// Mitsubishi GX Works2 project: Cascade3_V4   PLC: FX3G

TYPE PUMP : STRUCT
  Blocked : BOOL;
  Start : BOOL;
  Evailable : BOOL;
END_STRUCT END_TYPE

TYPE BURNER : STRUCT
  Manual : BOOL;
  Auto : BOOL;
  Stage1 : BOOL;
  Stage2 : BOOL;
  Pressure : INT;
  Temperature : INT;
  Power : BOOL;
  Work : BOOL;
  ManualSecond : BOOL;  (* Назначить горелку на вторую ступень *)
  Error : BOOL;
  Enable : BOOL;
END_STRUCT END_TYPE

// global labels: IO
VAR_GLOBAL
  AI_T_Heater1 AT D0 : INT;  (* Температура котла №1 с модуля АЦП (R23700), °C x10 *)
  AI_T_Heater2 AT D1 : INT;  (* Температура котла №2 с модуля АЦП (R23701), °C x10 *)
  AI_T_Heater3 AT D2 : INT;  (* Температура котла №3 с модуля АЦП (R23702), °C x10 *)
  AI_T_Colector AT D3 : INT;  (* Температура обратки с коллектора (R23703), °C x10 *)
  AI_T_SOFrom AT D4 : INT;  (* Температура обратки отопления (R23704), °C x10 *)
  AI_T_SOTo AT D5 : INT;  (* Температура подачи отопления (R23705), °C x10 *)
  AI_T_GVSTo AT D6 : INT;  (* Температура подачи на теплообменник ГВС (R23706), °C x10 *)
  AI_T_GVSFrom AT D7 : INT;  (* Температура обратки с теплообменника ГВС (R23707), °C x10 *)
  AI_T_Gaz AT D8 : INT;  (* Температура газа (R23709), °C x10 *)
  AI_T_Weather AT D9 : INT;  (* Температура наружного воздуха (R23708), °C x10 *)
  AI_P1 AT D10 : INT;  (* Давление в котле №1 с датчика, в десятых долях (шкала задаётся в Max_P1) *)
  AI_P2 AT D11 : INT;  (* Давление в котле №2 с датчика, в десятых долях (шкала задаётся в Max_P2) *)
  AI_P3 AT D12 : INT;  (* Давление в котле №3 с датчика, в десятых долях (шкала задаётся в Max_P3) *)
  AI_P_SOTo AT D13 : INT;  (* Давление подачи отопления с датчика, в десятых долях (шкала задаётся в Max_P_SOTo) *)
  AI_P_SOFrom AT D14 : INT;  (* Давление обратки отопления с датчика, в десятых долях (шкала задаётся в Max_P_SOFrom) *)
  AI_P_GVSTo AT D15 : INT;  (* Давление подачи на теплообменник с датчика, в десятых долях (шкала задаётся в Max_P_GVSTo) *)
  AI_P_GVSFrom AT D16 : INT;  (* Давление обратки с теплообменника с датчика, в десятых долях (шкала задаётся в Max_P_GVSFrom) *)
  AI_P_Set AT D17 : INT;  (* Давление в системе (подпитка), в десятых долях. D35 занят, поэтому D17 *)
  AI_P_GAZ AT D18 : INT;  (* Давление газа с датчика (D8032), в десятых долях *)
  DI_EKM AT X000 : BOOL;  (* Реле давления (ЭКМ): контакт разомкнут — авария 26 *)
  DI_ES AT X001 : BOOL;  (* Кнопка аварийного отключения: снимает gxStart, авария 27 *)
  DI_RKF AT X010 : BOOL;  (* Реле контроля фаз: контакт разомкнут — авария 28 *)
  DI_BurnAlarm1 AT X002 : BOOL;  (* Сухой контакт «авария горелки №1» *)
  DI_BurnAlarm2 AT X003 : BOOL;  (* Сухой контакт «авария горелки №2» *)
  DI_BurnAlarm3 AT X004 : BOOL;  (* Сухой контакт «авария горелки №3» *)
  DI_BurnWork1 AT X005 : BOOL;  (* Сухой контакт «горелка №1 в работе» *)
  DI_BurnWork2 AT X006 : BOOL;  (* Сухой контакт «горелка №2 в работе» *)
  DI_BurnWork3 AT X007 : BOOL;  (* Сухой контакт «горелка №3 в работе» *)
  DI_Pump1_T1 AT X011 : BOOL;  (* Обратная связь: насос №1 контура Т1 работает *)
  DI_Pump2_T1 AT X012 : BOOL;  (* Обратная связь: насос №2 контура Т1 работает *)
  DI_Pump1_T1_2 AT X013 : BOOL;  (* Обратная связь: насос №1 контура Т1.2 работает *)
  DI_Pump2_T1_2 AT X020 : BOOL;  (* Обратная связь: насос №2 контура Т1.2 работает *)
  DI_Pump1_T3 AT X021 : BOOL;  (* Обратная связь: насос №1 контура Т3 работает *)
  DI_Pump2_T3 AT X022 : BOOL;  (* Обратная связь: насос №2 контура Т3 работает *)
  DI_Pump1 AT X023 : BOOL;  (* Обратная связь: насос циркуляции №1 малого контура работает *)
  DI_Pump2 AT X024 : BOOL;  (* Обратная связь: насос циркуляции №2 малого контура работает *)
  DI_Pump3 AT X025 : BOOL;  (* Обратная связь: насос циркуляции №3 малого контура работает *)
  DI_AlarmReset AT X030 : BOOL;  (* Внешняя кнопка сброса аварий и сирены *)
  DI_BurnTherm1 AT X035 : BOOL;  (* Термозащита котла №1: нормально замкнутый контакт, нет цепи — авария *)
  DI_BurnTherm2 AT X036 : BOOL;  (* Термозащита котла №2: нормально замкнутый контакт, нет цепи — авария *)
  DI_BurnTherm3 AT X037 : BOOL;  (* Термозащита котла №3: нормально замкнутый контакт, нет цепи — авария *)
  DO_Burn1Power AT Y035 : BOOL;  (* Разрешение работы (питание) горелки №1: без него ступени не включаются *)
  DO_Burn1Stage1 AT Y000 : BOOL;  (* Горелка №1: включить ступень 1 *)
  DO_Burn1Stage2 AT Y001 : BOOL;  (* Горелка №1: включить ступень 2 *)
  DO_Burn2Power AT Y036 : BOOL;  (* Разрешение работы (питание) горелки №2: без него ступени не включаются *)
  DO_Burn2Stage1 AT Y002 : BOOL;  (* Горелка №2: включить ступень 1 *)
  DO_Burn2Stage2 AT Y003 : BOOL;  (* Горелка №2: включить ступень 2 *)
  DO_Burn3Power AT Y037 : BOOL;  (* Разрешение работы (питание) горелки №3: без него ступени не включаются *)
  DO_Burn3Stage1 AT Y004 : BOOL;  (* Горелка №3: включить ступень 1 *)
  DO_Burn3Stage2 AT Y005 : BOOL;  (* Горелка №3: включить ступень 2 *)
  DO_ValveFill AT Y006 : BOOL;  (* Клапан набора воды (подпитка) *)
  DO_AlarmBuzzer AT Y007 : BOOL;  (* Сирена: звуковая сигнализация аварии *)
  DO_AlarmLight AT Y010 : BOOL;  (* Лампа аварии *)
  DO_Pump1_T1 AT Y020 : BOOL;  (* Включить насос №1 контура Т1 *)
  DO_Pump2_T1 AT Y021 : BOOL;  (* Включить насос №2 контура Т1 *)
  DO_Pump1_T1_2 AT Y022 : BOOL;  (* Включить насос №1 контура Т1.2 *)
  DO_Pump2_T1_2 AT Y023 : BOOL;  (* Включить насос №2 контура Т1.2 *)
  DO_Pump1_T3 AT Y024 : BOOL;  (* Включить насос №1 контура Т3 *)
  DO_Pump2_T3 AT Y025 : BOOL;  (* Включить насос №2 контура Т3 *)
  DO_Pump1 AT Y026 : BOOL;  (* Включить насос циркуляции №1 малого контура *)
  DO_Pump2 AT Y027 : BOOL;  (* Включить насос циркуляции №2 малого контура *)
  DO_Pump3 AT Y030 : BOOL;  (* Включить насос циркуляции №3 малого контура *)
  DO_3wayOpen AT Y033 : BOOL;  (* 3-ходовой клапан: открыть *)
  DO_3wayClose AT Y034 : BOOL;  (* 3-ходовой клапан: закрыть *)
END_VAR

// global labels: GVL
VAR_GLOBAL
  arBurners : ARRAY [0..2] OF BURNER;  (* (Set M500) Состояние трёх котлов (структура BURNER): включён в авто, ступень 1, ступень 2, авария, ручной режим *)
END_VAR
VAR_GLOBAL CONSTANT
  c_HEATERS : INT := 3;  (* Количество котлов в каскаде *)
  c_HEATERS_IDX : INT := 2;  (* Индекс последнего котла в массиве (c_HEATERS - 1) *)
  c_AM_ALARMS_NUM : INT := 54;  (* Верхняя граница массива аварий: используются номера 0…45 (46 штук). Максимум 127 *)
END_VAR
VAR_GLOBAL
  AM_ALARMS : ARRAY [0..54] OF ST_AM_ALARM;  (* Массив аварий менеджера тревог. Граница 45 должна совпадать с c_AM_ALARMS_NUM. Состояние: AM_ALARMS[i].Alarm *)
  gxStart AT M400 : BOOL;  (* Пуск/останов каскада с панели (1 = работа). Снимается кнопкой X001 и авариями *)
  gxErrorReset AT M401 : BOOL;  (* Сброс всех аварий (1 = сбросить). В шаге 0 выставляется программой автоматически *)
  gxHasalarm AT M402 : BOOL;  (* Есть хотя бы одна активная авария. Формируется блоком FB_AM_HAS_ALARMS, используется для лампы и панели *)
  gxNoSettings AT M403 : BOOL;  (* Не заданы уставки или коэффициенты ПИД (R503 = 0). Пуск запрещён, авария 30 *)
  gxResetAlarm AT M404 : BOOL;  (* Кнопка «Сброс сигнализации» на панели: снимает сирену и лампу *)
  gxFillManual AT M405 : BOOL;  (* Ручной режим подпитки: клапан набора воды открыт, пока флаг включён *)
  gxFillAuto AT M406 : BOOL;  (* Автоматическая подпитка по давлению в системе (SV_PresFilStart / SV_PresFilStop) *)
  gxResetWHT1 AT M407 : BOOL;  (* Сброс моточасов котла №1 (giHeater1Hours) *)
  gxResetWHT2 AT M408 : BOOL;  (* Сброс моточасов котла №2 (giHeater2Hours) *)
  gxResetWHT3 AT M409 : BOOL;  (* Сброс моточасов котла №3 (giHeater3Hours) *)
  gxPIDAT AT M410 : BOOL;  (* Запуск автонастройки ПИД каскада (блок параметров R500…R528). Сбрасывается сама по завершении *)
  gxPIDATLimitCycle AT M411 : BOOL;  (* Ограничение числа циклов автонастройки ПИД каскада: 0 — не больше 50, 1 — не больше 114 *)
  gxEnablePump1 AT M412 : BOOL;  (* Разрешение насоса циркуляции №1 малого контура (1 = участвует в работе) *)
  gxEnablePump2 AT M413 : BOOL;  (* Разрешение насоса циркуляции №2 малого контура (1 = участвует в работе) *)
  gxEnablePump3 AT M415 : BOOL;  (* Разрешение насоса циркуляции №3 малого контура (1 = участвует в работе). M414 пропущен — так привязано на панели *)
  gxManualPump1 AT M416 : BOOL;  (* Ручной пуск насоса циркуляции №1 малого контура (нужно ещё разрешение gxEnablePump1) *)
  gxManualPump2 AT M417 : BOOL;  (* Ручной пуск насоса циркуляции №2 малого контура (нужно ещё разрешение gxEnablePump2) *)
  gxManualPump3 AT M418 : BOOL;  (* Ручной пуск насоса циркуляции №3 малого контура (нужно ещё разрешение gxEnablePump3) *)
  gx3WayCloseWhenOff AT M419 : BOOL;  (* Закрывать 3-ходовой клапан при останове каскада (1 = закрывать) *)
  gxPID3WayAT AT M420 : BOOL;  (* Запуск автонастройки ПИД 3-ходового клапана (блок параметров R600…R628) *)
  gxPID3WayATLimitCycle AT M421 : BOOL;  (* Ограничение числа циклов автонастройки ПИД 3-ходового клапана: 0 — не больше 50, 1 — не больше 114 *)
  gxPump1_T1_Enable AT M422 : BOOL;  (* Разрешение насоса №1 контура Т1 (1 = участвует в каскаде, 0 = заблокирован) *)
  gxPump2_T1_Enable AT M423 : BOOL;  (* Разрешение насоса №2 контура Т1 (1 = участвует в каскаде, 0 = заблокирован) *)
  gxPump1_T1_2_Enable AT M424 : BOOL;  (* Разрешение насоса №1 контура Т1.2 (1 = участвует в каскаде, 0 = заблокирован) *)
  gxPump2_T1_2_Enable AT M425 : BOOL;  (* Разрешение насоса №2 контура Т1.2 (1 = участвует в каскаде, 0 = заблокирован) *)
  gxPump1_T3_Enable AT M426 : BOOL;  (* Разрешение насоса №1 контура Т3 (1 = участвует в каскаде, 0 = заблокирован) *)
  gxPump2_T3_Enable AT M427 : BOOL;  (* Разрешение насоса №2 контура Т3 (1 = участвует в каскаде, 0 = заблокирован) *)
  gxPump1_T1_Manual AT M428 : BOOL;  (* Ручной пуск насоса №1 контура Т1 *)
  gxPump2_T1_Manual AT M429 : BOOL;  (* Ручной пуск насоса №2 контура Т1 *)
  gxPump1_T1_2_Manual AT M430 : BOOL;  (* Ручной пуск насоса №1 контура Т1.2 *)
  gxPump2_T1_2_Manual AT M431 : BOOL;  (* Ручной пуск насоса №2 контура Т1.2 *)
  gxPump1_T3_Manual AT M432 : BOOL;  (* Ручной пуск насоса №1 контура Т3 *)
  gxPump2_T3_Manual AT M433 : BOOL;  (* Ручной пуск насоса №2 контура Т3 *)
  gxPump1_T1_WHReset AT M434 : BOOL;  (* Сброс моточасов насоса №1 контура Т1 *)
  gxPump2_T1_WHReset AT M435 : BOOL;  (* Сброс моточасов насоса №2 контура Т1 *)
  gxPump1_T1_2_WHReset AT M436 : BOOL;  (* Сброс моточасов насоса №1 контура Т1.2 *)
  gxPump2_T1_2_WHReset AT M437 : BOOL;  (* Сброс моточасов насоса №2 контура Т1.2 *)
  gxPump1_T3_WHReset AT M438 : BOOL;  (* Сброс моточасов насоса №1 контура Т3 *)
  gxPump2_T3_WHReset AT M439 : BOOL;  (* Сброс моточасов насоса №2 контура Т3 *)
  gxPump1_WHReset AT M440 : BOOL;  (* Сброс моточасов насоса циркуляции №1 малого контура *)
  gxPump2_WHReset AT M441 : BOOL;  (* Сброс моточасов насоса циркуляции №2 малого контура *)
  gxPump3_WHReset AT M442 : BOOL;  (* Сброс моточасов насоса циркуляции №3 малого контура *)
  gx3WayEnable AT M443 : BOOL;  (* Разрешение работы 3-ходового клапана (1 = регулирует, 0 = стоит) *)
  gx3WayManual AT M444 : BOOL;  (* Ручной режим 3-ходового клапана: положение берётся из SV_3WayManualTask, ПИД отключён *)
  gxWHOvfHeater1 AT M450 : BOOL;  (* Переполнение счётчика моточасов котла №1 (выход HOUR). 1 — счётчик переполнен, нужно сбросить *)
  gxWHOvfHeater2 AT M451 : BOOL;  (* Переполнение счётчика моточасов котла №2 (выход HOUR). 1 — счётчик переполнен, нужно сбросить *)
  gxWHOvfHeater3 AT M452 : BOOL;  (* Переполнение счётчика моточасов котла №3 (выход HOUR). 1 — счётчик переполнен, нужно сбросить *)
  gxWHOvfPump1_T1 AT M453 : BOOL;  (* Переполнение счётчика моточасов насоса №1 контура Т1 (выход HOUR) *)
  gxWHOvfPump2_T1 AT M454 : BOOL;  (* Переполнение счётчика моточасов насоса №2 контура Т1 (выход HOUR) *)
  gxWHOvfPump1_T1_2 AT M455 : BOOL;  (* Переполнение счётчика моточасов насоса №1 контура Т1.2 (выход HOUR) *)
  gxWHOvfPump2_T1_2 AT M456 : BOOL;  (* Переполнение счётчика моточасов насоса №2 контура Т1.2 (выход HOUR) *)
  gxWHOvfPump1_T3 AT M457 : BOOL;  (* Переполнение счётчика моточасов насоса №1 контура Т3 (выход HOUR) *)
  gxWHOvfPump2_T3 AT M458 : BOOL;  (* Переполнение счётчика моточасов насоса №2 контура Т3 (выход HOUR) *)
  gxWHOvfPump1 AT M459 : BOOL;  (* Переполнение счётчика моточасов насоса циркуляции №1 (выход HOUR) *)
  gxWHOvfPump2 AT M460 : BOOL;  (* Переполнение счётчика моточасов насоса циркуляции №2 (выход HOUR) *)
  gxWHOvfPump3 AT M461 : BOOL;  (* Переполнение счётчика моточасов насоса циркуляции №3 (выход HOUR) *)
  giPIDTask AT D500 : INT;  (* Выход ПИД каскада: задание в ступенях мощности (0…6). Из него считается, сколько котлов и ступеней включить *)
  giTSV AT D501 : INT;  (* Текущее задание температуры теплоносителя: по кривой погодозависимости или SV_TWater1, если на улице тепло *)
  giAvailableStages AT D502 : INT;  (* Сколько ступеней доступно автоматике: по 2 на каждый котёл в авто без аварий *)
  giWorkStages AT D503 : INT;  (* Сколько ступеней включено сейчас в авторежиме *)
  giPID3WayTask AT D504 : INT;  (* Выход ПИД 3-ходового клапана: положение 0…1000 (0.0…100.0 %, 0 — закрыт, 1000 — открыт). Диапазон задан R622 = 1000 *)
  SV_3WayTempGVS AT D510 : INT;  (* Уставка температуры ГВС на выходе теплообменника, °C *)
  SV_MaxTemperatureHeater AT D511 : INT;  (* Максимальная температура котла, °C. Выше — авария перегрева *)
  SV_TLimit AT D512 : INT;  (* Допустимое превышение задания, °C: котёл отключается при температуре выше задания на эту величину *)
  SV_HowOftenToCheck AT D513 : INT;  (* Как часто проверять каскад (добавлять или убирать ступени), секунд *)
  SV_MaxPressure AT D514 : INT;  (* Максимальное давление в котле (авария). В тех же единицах, что и показания датчика *)
  SV_MinPressure AT D515 : INT;  (* Минимальное давление в котле (авария) *)
  SV_PresFilStart AT D516 : INT;  (* Давление в системе, при котором начинается подпитка *)
  SV_PresFilStop AT D517 : INT;  (* Давление в системе, при котором подпитка заканчивается *)
  SV_GasMinPressure AT D518 : INT;  (* Минимальное давление газа. Ниже — авария 24 и блокировка каскада *)
  SV_SetMinPressure AT D519 : INT;  (* Минимальное давление в системе. Ниже — авария 25 и запрет циркуляционных насосов *)
  SV_MaxFillTime AT D520 : INT;  (* Максимальное время набора воды, секунд. Дольше — авария 34 *)
  SV_TimeinWork AT D521 : INT;  (* Резерв: в программе не используется (осталось от старой версии), выводится только на панель *)
  SV_3WayDelta AT D522 : INT;  (* Зона нечувствительности 3-ходового клапана в единицах положения 0…1000 (50 = 5.0 %); в ручном режиме принудительно равна 0 *)
  SV_3WayTotalTime AT D523 : INT;  (* Полное время хода 3-ходового клапана, секунд *)
  SV_3WayLuftTime AT D524 : INT;  (* Время люфта (мёртвого хода) 3-ходового клапана, миллисекунд *)
  SV_3WayTempGVSDelta AT D525 : INT;  (* Гистерезис по ГВС, °C: ПИД работает, пока температура ниже уставки на эту величину *)
  SV_3WayManualTask AT D526 : INT;  (* Задание положения 3-ходового клапана в ручном режиме, 0…1000 (0.1 % за единицу) — та же шкала, что у выхода ПИД *)
  SV_3WayMaxTemperature AT D527 : INT;  (* Максимальная температура ГВС, °C. Выше — авария 35 *)
  SV_MaxTemperatureColector AT D528 : INT;  (* Максимальная температура коллектора, °C. Выше — авария 32 и отключение ПИД каскада *)
  SV_StageHyst AT D583 : INT;  (* % x10 с панели (50 = 5.0 %). Зона нечувствительности добавления ступени: насколько выход ПИД (0…600 = 0…100 %) должен превысить границу следующей ступени, чтобы включилась ещё одна ступень. Убираются ступени без задержки. ПЛК пересчитывает проценты в единицы ПИД: iHyst = значение * 6 / 10 *)
  giHeater1Hours AT D560 : ARRAY [0..1] OF INT;  (* Наработка котла №1, моточасы (массив из 2 слов для счётчика HOUR) *)
  giHeater2Hours AT D562 : ARRAY [0..1] OF INT;  (* Наработка котла №2, моточасы (массив из 2 слов для счётчика HOUR) *)
  giHeater3Hours AT D564 : ARRAY [0..1] OF INT;  (* Наработка котла №3, моточасы (массив из 2 слов для счётчика HOUR) *)
  T1_State AT D566 : INT;  (* Состояние котла №1 для панели: 0 — не разрешён, 1 — разрешён и стоит, 2 — ступень 1, 3 — ступень 2 *)
  T2_State AT D567 : INT;  (* Состояние котла №2 для панели: 0 — не разрешён, 1 — разрешён и стоит, 2 — ступень 1, 3 — ступень 2 *)
  T3_State AT D568 : INT;  (* Состояние котла №3 для панели: 0 — не разрешён, 1 — разрешён и стоит, 2 — ступень 1, 3 — ступень 2 *)
  Pump1_T1_State AT D569 : INT;  (* Состояние насоса №1 контура Т1 для панели: 0 — стоит, 1 — работает, 2 — авария, 4 — заблокирован *)
  Pump2_T1_State AT D570 : INT;  (* Состояние насоса №2 контура Т1 для панели: 0 — стоит, 1 — работает, 2 — авария, 4 — заблокирован *)
  Pump1_T1_2_State AT D571 : INT;  (* Состояние насоса №1 контура Т1.2 для панели: 0 — стоит, 1 — работает, 2 — авария, 4 — заблокирован *)
  Pump2_T1_2_State AT D572 : INT;  (* Состояние насоса №2 контура Т1.2 для панели: 0 — стоит, 1 — работает, 2 — авария, 4 — заблокирован *)
  Pump1_T3_State AT D573 : INT;  (* Состояние насоса №1 контура Т3 для панели: 0 — стоит, 1 — работает, 2 — авария, 4 — заблокирован *)
  Pump2_T3_State AT D574 : INT;  (* Состояние насоса №2 контура Т3 для панели: 0 — стоит, 1 — работает, 2 — авария, 4 — заблокирован *)
  Pump1_State AT D575 : INT;  (* Состояние насоса циркуляции №1 для панели: 0 — стоит, 1 — работает, 2 — авария, 4 — заблокирован *)
  Pump2_State AT D576 : INT;  (* Состояние насоса циркуляции №2 для панели: 0 — стоит, 1 — работает, 2 — авария, 4 — заблокирован *)
  Pump3_State AT D577 : INT;  (* Состояние насоса циркуляции №3 для панели: 0 — стоит, 1 — работает, 2 — авария, 4 — заблокирован *)
  Pump1_T1_WH AT D600 : ARRAY [0..1] OF INT;  (* Моточасы насоса №1 контура Т1 (2 слова, счётчик HOUR). Область D600…D617 не пересекается с состояниями *)
  Pump2_T1_WH AT D602 : ARRAY [0..1] OF INT;  (* Моточасы насоса №2 контура Т1 (2 слова, счётчик HOUR). Область D600…D617 не пересекается с состояниями *)
  Pump1_T1_2_WH AT D604 : ARRAY [0..1] OF INT;  (* Моточасы насоса №1 контура Т1.2 (2 слова, счётчик HOUR). Область D600…D617 не пересекается с состояниями *)
  Pump2_T1_2_WH AT D606 : ARRAY [0..1] OF INT;  (* Моточасы насоса №2 контура Т1.2 (2 слова, счётчик HOUR). Область D600…D617 не пересекается с состояниями *)
  Pump1_T3_WH AT D608 : ARRAY [0..1] OF INT;  (* Моточасы насоса №1 контура Т3 (2 слова, счётчик HOUR). Область D600…D617 не пересекается с состояниями *)
  Pump2_T3_WH AT D610 : ARRAY [0..1] OF INT;  (* Моточасы насоса №2 контура Т3 (2 слова, счётчик HOUR). Область D600…D617 не пересекается с состояниями *)
  Pump1_WH AT D612 : ARRAY [0..1] OF INT;  (* Моточасы насоса циркуляции №1 (2 слова, счётчик HOUR). Область D600…D617 не пересекается с состояниями *)
  Pump2_WH AT D614 : ARRAY [0..1] OF INT;  (* Моточасы насоса циркуляции №2 (2 слова, счётчик HOUR). Область D600…D617 не пересекается с состояниями *)
  Pump3_WH AT D616 : ARRAY [0..1] OF INT;  (* Моточасы насоса циркуляции №3 (2 слова, счётчик HOUR). Область D600…D617 не пересекается с состояниями *)
  SV_TWeather1 AT D530 : INT;  (* Кривая погодозависимости, точка 1: температура на улице, °C *)
  SV_TWater1 AT D531 : INT;  (* Кривая погодозависимости, точка 1: температура подачи в систему, °C *)
  SV_TWeather2 AT D532 : INT;  (* Кривая погодозависимости, точка 2: температура на улице, °C *)
  SV_TWater2 AT D533 : INT;  (* Кривая погодозависимости, точка 2: температура подачи в систему, °C *)
  SV_TWeather3 AT D534 : INT;  (* Кривая погодозависимости, точка 3: температура на улице, °C *)
  SV_TWater3 AT D535 : INT;  (* Кривая погодозависимости, точка 3: температура подачи в систему, °C *)
  SV_TWeather4 AT D536 : INT;  (* Кривая погодозависимости, точка 4: температура на улице, °C *)
  SV_TWater4 AT D537 : INT;  (* Кривая погодозависимости, точка 4: температура подачи в систему, °C *)
  Cor_T_Heater1 AT D540 : INT;  (* Поправка датчика температуры котла №1: прибавляется к показанию, °C x10 *)
  Cor_T_Heater2 AT D541 : INT;  (* Поправка датчика температуры котла №2: прибавляется к показанию, °C x10 *)
  Cor_T_Heater3 AT D542 : INT;  (* Поправка датчика температуры котла №3: прибавляется к показанию, °C x10 *)
  Cor_T_Colector AT D543 : INT;  (* Поправка датчика температуры коллектора: прибавляется к показанию, °C x10 *)
  Cor_T_SOFrom AT D544 : INT;  (* Поправка датчика температуры обратки отопления: прибавляется к показанию, °C x10 *)
  Cor_T_SOTo AT D545 : INT;  (* Поправка датчика температуры подачи отопления: прибавляется к показанию, °C x10 *)
  Cor_T_GVSTo AT D546 : INT;  (* Поправка датчика температуры подачи на теплообменник ГВС: прибавляется к показанию, °C x10 *)
  Cor_T_GVSFrom AT D547 : INT;  (* Поправка датчика температуры обратки с теплообменника ГВС: прибавляется к показанию, °C x10 *)
  Cor_T_Gaz AT D548 : INT;  (* Поправка датчика температуры датчика газа: прибавляется к показанию, °C x10 *)
  Cor_T_Weather AT D549 : INT;  (* Поправка датчика температуры датчика наружной температуры: прибавляется к показанию, °C x10 *)
  Max_P1 AT D550 : INT;  (* Верхний предел шкалы датчика давления котла №1, в десятых долях (160 = 16.0). 0 — не задан *)
  Max_P2 AT D551 : INT;  (* Верхний предел шкалы датчика давления котла №2, в десятых долях (160 = 16.0). 0 — не задан *)
  Max_P3 AT D552 : INT;  (* Верхний предел шкалы датчика давления котла №3, в десятых долях (160 = 16.0). 0 — не задан *)
  Max_P_SOTo AT D553 : INT;  (* Верхний предел шкалы датчика давления подачи отопления, в десятых долях (160 = 16.0). 0 — не задан *)
  Max_P_SOFrom AT D554 : INT;  (* Верхний предел шкалы датчика давления обратки отопления, в десятых долях (160 = 16.0). 0 — не задан *)
  Max_P_GVSTo AT D555 : INT;  (* Верхний предел шкалы датчика давления подачи на теплообменник, в десятых долях (160 = 16.0). 0 — не задан *)
  Max_P_GVSFrom AT D556 : INT;  (* Верхний предел шкалы датчика давления обратки с теплообменника, в десятых долях (160 = 16.0). 0 — не задан *)
  Max_P_Set AT D557 : INT;  (* Верхний предел шкалы датчика давления в системе, в десятых долях (160 = 16.0). 0 — не задан *)
  Max_P_GAZ AT D558 : INT;  (* Верхний предел шкалы датчика давления газа, в десятых долях (160 = 16.0). 0 — не задан *)
  FAI_T_Heater1 AT D20 : REAL;  (* Температура котла №1, °C в реальных единицах (для панели и графиков) *)
  FAI_T_Heater2 AT D22 : REAL;  (* Температура котла №2, °C в реальных единицах (для панели и графиков) *)
  FAI_T_Heater3 AT D24 : REAL;  (* Температура котла №3, °C в реальных единицах (для панели и графиков) *)
  FAI_T_Colector AT D26 : REAL;  (* Температура обратки с коллектора, °C в реальных единицах (для панели и графиков) *)
  FAI_T_SOFrom AT D28 : REAL;  (* Температура обратки отопления, °C в реальных единицах (для панели и графиков) *)
  FAI_T_SOTo AT D30 : REAL;  (* Температура подачи отопления, °C в реальных единицах (для панели и графиков) *)
  FAI_T_GVSTo AT D32 : REAL;  (* Температура подачи на теплообменник ГВС, °C в реальных единицах (для панели и графиков) *)
  FAI_T_GVSFrom AT D34 : REAL;  (* Температура обратки с теплообменника ГВС, °C в реальных единицах (для панели и графиков) *)
  FAI_T_Gaz AT D36 : REAL;  (* Температура газа, °C в реальных единицах (для панели и графиков) *)
  FAI_T_Weather AT D38 : REAL;  (* Температура наружного воздуха, °C в реальных единицах (для панели и графиков) *)
  FAI_P1 AT D40 : REAL;  (* Давление в котле №1 в реальных единицах (для панели и графиков) *)
  FAI_P2 AT D42 : REAL;  (* Давление в котле №2 в реальных единицах (для панели и графиков) *)
  FAI_P3 AT D44 : REAL;  (* Давление в котле №3 в реальных единицах (для панели и графиков) *)
  FAI_P_SOTo AT D46 : REAL;  (* Давление подачи отопления в реальных единицах (для панели и графиков) *)
  FAI_P_SOFrom AT D48 : REAL;  (* Давление обратки отопления в реальных единицах (для панели и графиков) *)
  FAI_P_GVSTo AT D50 : REAL;  (* Давление подачи на теплообменник в реальных единицах (для панели и графиков) *)
  FAI_P_GVSFrom AT D52 : REAL;  (* Давление обратки с теплообменника в реальных единицах (для панели и графиков) *)
  FAI_P_Set AT D54 : REAL;  (* Давление в системе в реальных единицах (для панели и графиков) *)
  FAI_P_GAZ AT D56 : REAL;  (* Давление газа в реальных единицах (для панели и графиков) *)
END_VAR

// task Task_01 (event TRUE, interval 0, priority 31): POU_01
// task PROCESS (event FALSE, interval T#50ms, priority 2): PROCESS
// task INIT (event M8002, interval 0, priority 1): INIT
// task TCO (event I750, interval 0, priority 25): PRG_TCO_TICKER_50
// user libraries (not included): AlarmManager, TimeControl, Utils

PROGRAM POU_01
VAR
  fbAmBlock : FB_AM_IS_BLOCK;
  fbCirculation : Circulation;
  fbValve : FB_VALVE_3P;
  fbPumpsSO : PUMPS;
  fbPumpsToTO : PUMPS;
  fbPumpsFromTO : PUMPS;
  xIsError : BOOL;
  xPIDWork : BOOL;
  xPID3WayWork : BOOL;
  iStep : INT;  (* Текущий шаг *)
  iCount : INT;
  iCountStages : INT;  (* Всего на данный момент задействовано степеней по 2 на горелку *)
  iReverced : INT;  (* Индекс котла в обратном порядке от 5 до 0 *)
  iShifted : INT;  (* Индекс котла с учетом сдвига *)
  iShifter : INT;  (* На сколько нужно сделать сдвиг *)
  iToSubtract : INT;  (* Сколько степеней нужно убавить *)
  iStepSize : INT;  (* Цена одной ступени в процентах выхода ПИД (R522 / число доступных ступеней) *)
  iHyst : INT;  (* Зона нечувствительности добавления ступени в единицах выхода ПИД (из «Дельта %» с панели: 50 = 5.0 % = 30 единиц) *)
  iAddLimit : INT;  (* Порог выхода ПИД, при котором добавляется следующая ступень (граница ступени + iHyst) *)
  iPIDMax : INT;  (* Верхний предел выхода ПИД каскада (копия R522 из блока параметров R500..R528), 600 = 100 % *)
  iToAdd : INT;  (* Скольо степеней нужно добавить *)
END_VAR
EI(TRUE);

(* Шаги селектора ступеней (iStep):
   0 - инициализация, 1 - промежуточный, 2 - выключить все горелки,
   3 - ожидание пуска, 4 - расчёт числа ступеней по заданию ПИД,
   5 - работа (ждём TC13 или отказа котла) *)

fbAmBlock(iProcessNum := 10, iSeverity := c_AM_ERROR);

(* stop s knopki *)
RST(NOT DI_ES , gxStart);

(* Если общий блок то выключаем все горелки *)
MOV(fbAmBlock.Q AND NOT (iStep = 3), 2, iStep);
MOV(MEF(gxStart), 2, iStep);

(* Как часто заходить в селектор. TC13 - таймер с базой 100 мс,
   SV_HowOftenToCheck задаётся с панели в СЕКУНДАХ, поэтому * 10 *)
OUT_T(iStep = 5, TC13, SV_HowOftenToCheck * 10);

(* PID for heating *)
xPIDWork :=
    (iStep = 4 OR iStep = 5)
    AND (AI_T_Colector < (giTSV + SV_TLimit))
    (* Обрыв датчика коллектора (авария 39): без обратной связи ПИД ушёл бы
       на 100 %, поэтому регулятор снимается и задание каскада обнуляется *)
    AND NOT AM_ALARMS[39].Alarm
    AND NOT fbAmBlock.Q;
(* Если включена автонастройка ПИД то активируем *)
MOVP(
    xPIDWork AND gxPIDAT,
    SEL(gxPIDATLimitCycle, 2#0000_0000_0011_0001, 2#0000_0000_0111_0001),
    R501
);
(* Если начали Автонастроку то отключаем этот параметр *)
RST(xPIDWork AND gxPIDAT, gxPIDAT);

PID(xPIDWork, giTSV, AI_T_Colector, R500, giPIDTask);
(* Если регулятор не работает, задание на каскад = 0 (все ступени выкл.) *)
MOV(NOT xPIDWork, 0, giPIDTask);

CASE iStep OF
0: (* Init *)
    gxStart := 0;
    gxErrorReset := TRUE;
    iStep := 1;
1:
    iStep := 2;
2: (* Сброс при блокировке работы *)
    FOR iCount := 0 TO c_HEATERS_IDX DO
        arBurners[iCount].Power := FALSE;
        arBurners[iCount].Stage1 := FALSE;
        arBurners[iCount].Stage2 := FALSE;
    END_FOR;

    iStep := 3;

3: (* idle *)
    IF gxStart AND NOT fbAmBlock.Q THEN
        (* Смещаем индекс основной котел 0-5 для 6ти котолов *)
        (* TODO: смещение раз в неделю добавить *)
        iShifter := F_INCN(TRUE, iShifter, c_HEATERS_IDX);
        iStep := 4;
    END_IF;

4: (* select *)
    iCountStages := 0; (* Текущие ступени в авто *)
    giAvailableStages := 0; (* Всего доступно ступеней в авто *)
    FOR iCount := 0 TO c_HEATERS_IDX DO
        arBurners[iCount].Power := (
            arBurners[iCount].Auto OR arBurners[iCount].Manual
        ) AND NOT arBurners[iCount].Error AND arBurners[iCount].Enable;

        IF arBurners[iCount].Manual AND arBurners[iCount].Power THEN
            (* Когда включаем в ручно, ступень тоже в ручном устанавливается *)
            arBurners[iCount].Stage1 := TRUE;
            arBurners[iCount].Stage2 := arBurners[iCount].ManualSecond;
        END_IF;

        IF arBurners[iCount].Auto AND NOT arBurners[iCount].Error THEN
            (* Считаем сколько ступеней уже включено в авто режиме *)
            INC(arBurners[iCount].Stage1, iCountStages);
            INC(arBurners[iCount].Stage2, iCountStages);
            (* Считаем сколько ступеней вообще доступно для авто режима *)
            INC(arBurners[iCount].Power, giAvailableStages);
            INC(arBurners[iCount].Power, giAvailableStages);
        END_IF;
    END_FOR;

    (* Найти сколько еще нужно включить котлов
    R522 это максимальная задача ПИД регулятора *)
    (* Защита от деления на ноль: если нет ни одного котла в авто
       (все в ручном, в аварии или запрещены) или цена ступени нулевая,
       шаг не считаем. Через IF, а не SEL: ST вычисляет все аргументы
       функции, поэтому деление на 0 всё равно произошло бы *)
    (* R522 - верхний предел выхода ПИД из блока параметров R500..R528
       (600 = 100 %). Копируем в именованную переменную, чтобы ниже
       не было "магического" номера регистра *)
    iPIDMax := R522;
    iStepSize := 0;
    IF giAvailableStages > 0 THEN
        iStepSize := iPIDMax / giAvailableStages;
    END_IF;

    (* ДОБАВЛЕНИЕ: не больше одной ступени за период проверки, чтобы мощность
       росла плавно. Ступень включается только если ПИД вышел за границу
       следующей ступени на зону нечувствительности, иначе на самой границе ступень
       дёргалась бы каждый период. У последней доступной ступени гистерезис
       не применяется (порог ограничен R522), иначе она не включилась бы
       никогда *)
    (* «Дельта %» с панели приходит в процентах x10 (50 = 5.0 %), а выход ПИД
       и цена ступени считаются в единицах 0…600 (100 %). Поэтому проценты
       переводим: 1 % = 6 единиц -> 5.0 % (50) = 30 единиц *)
    iHyst := SV_StageHyst * 6 / 10;

    iToAdd := 0;
    IF iStepSize > 0 AND iCountStages < giAvailableStages THEN
        iAddLimit := ((iCountStages + 1) * iStepSize) + iHyst;
        IF iAddLimit > iPIDMax THEN
            iAddLimit := iPIDMax;
        END_IF;
        IF giPIDTask >= iAddLimit THEN
            iToAdd := 1;
        END_IF;
    END_IF;

    (* УБАВЛЕНИЕ: снимаем сразу столько ступеней, сколько требует ПИД.
       Снижение мощности не задерживается никогда - опасен перегрев *)
    iToSubtract := 0;
    IF iStepSize > 0 THEN
        iToSubtract := iCountStages - (giPIDTask / iStepSize);
        IF iToSubtract < 0 THEN
            iToSubtract := 0;
        END_IF;
    END_IF;

    IF iToAdd > 0 THEN
        FOR iCount := 0 TO c_HEATERS_IDX DO
            (* Смещаем индек для выравнивания моточасов *)
            iShifted := F_SHFT(iShifter, iCount, c_HEATERS_IDX);
            IF iToAdd > 0
                AND arBurners[iShifted].Auto
                AND arBurners[iShifted].Power
            THEN
                (* Не запущен *)
                IF NOT arBurners[iShifted].Stage1 THEN
                    arBurners[iShifted].Stage1 := TRUE;
                    arBurners[iShifted].Stage2 := iToAdd > 1;
                    SUB_E(TRUE, iToAdd, 1, iToAdd);
                    SUB_E(arBurners[iShifted].Stage2, iToAdd, 1, iToAdd);
                (* Запущен только на одну ступень *)
                ELSIF (arBurners[iShifted].Stage1 AND NOT arBurners[iShifted].Stage2) THEN
                    arBurners[iShifted].Stage2 := TRUE;
                    SUB_E(TRUE, iToAdd, 1, iToAdd);
                END_IF;
            END_IF;

            (* Закончить цикл если больше не нужно добавлять
            TODO: добавить что добавляем только по одному котлу раз в период *)
            IF iToAdd <= 0 THEN EXIT; END_IF;
        END_FOR;

    ELSIF iToSubtract > 0 THEN
        FOR iCount := 0 TO c_HEATERS_IDX DO
            (* Проходим массив начиная с конца в начало *)
            iReverced := REVERSE(iCount, c_HEATERS_IDX);
            (* Смещаем индек для выравнивания моточасов *)
            iShifted := F_SHFT(iShifter, iReverced, c_HEATERS_IDX);
            IF iToSubtract > 0
                AND arBurners[iShifted].Auto
                AND arBurners[iShifted].Power
                AND arBurners[iShifted].Stage1
            THEN

                (* Запущен на две ступени *)
                IF arBurners[iShifted].Stage2 THEN
                    (* Выключаем если нужно понизить больше чем на 2 ступени *)
                    arBurners[iShifted].Stage1 := iToSubtract < 2;

                    (* Понижаем на одну степень как минимум *)
                    arBurners[iShifted].Stage2 := FALSE;
                    SUB_E(TRUE, iToSubtract, 1, iToSubtract);

                    (* Если выключили значит понизили на 2 ступени *)
                    SUB_E(NOT arBurners[iShifted].Stage1, iToSubtract, 1, iToSubtract);

                (* Запущен на одну ступень *)
                ELSE
                    arBurners[iShifted].Stage1 := FALSE;
                    SUB_E(TRUE, iToSubtract, 1, iToSubtract);
                END_IF;
            END_IF;

            (* Закончить цикл если больше не нужно выключать *)
            IF iToSubtract <= 0 THEN EXIT; END_IF;
        END_FOR;
    END_IF;

    iStep := 5;

5: (* work *)
    xIsError := FALSE;
    FOR iCount := 0 TO c_HEATERS_IDX DO
        IF (arBurners[iCount].Error OR NOT arBurners[iCount].Enable) AND arBurners[iCount].Power THEN
            arBurners[iCount].Manual := FALSE;
            arBurners[iCount].Power := FALSE;
            arBurners[iCount].Stage1 := FALSE;
            arBurners[iCount].Stage2 := FALSE;
            xIsError := TRUE;
        END_IF;
    END_FOR;
    (* Ecли откзал котел или время вышло, на селектор *)
    MOV(xIsError OR TS13, 4, iStep);
    MOV(NOT gxStart, 2, iStep); (* na 2 shag chtobi vse vikluchit *)
END_CASE;

FOR iCount := 0 TO c_HEATERS_IDX DO
    IF MEP(arBurners[iCount].Auto) THEN
        arBurners[iCount].Manual := FALSE;
        arBurners[iCount].ManualSecond := FALSE;
    END_IF;
    IF arBurners[iCount].Manual OR arBurners[iCount].ManualSecond THEN
        arBurners[iCount].Auto := FALSE;
    END_IF;
END_FOR;

(* 3way *)
xPID3WayWork := gx3WayEnable
    AND (iStep = 4 OR iStep = 5)
    AND (DO_Pump1_T1_2 OR DO_Pump2_T1_2)
    (* Обрыв датчика обратки ГВС (авария 43): ПИД клапана снимается,
       иначе он открыл бы клапан на 100 % по -199 C *)
    AND NOT AM_ALARMS[43].Alarm
    AND (AI_T_GVSFrom < SV_3WayTempGVS + SV_3WayTempGVSDelta);
MOVP(xPID3WayWork AND gxPID3WayAT, SEL(gxPID3WayATLimitCycle, 2#0000_0000_0011_0001, 2#0000_0000_0111_0001), R601);
RST(xPID3WayWork AND gxPID3WayAT, gxPID3WayAT);
PID(xPID3WayWork, SV_3WayTempGVS, AI_T_GVSFrom, R600, giPID3WayTask);
MOV(NOT xPID3WayWork, 0, giPID3WayTask);
RST(MEF(gx3WayEnable), gx3WayManual);
SET(gx3WayManual, gx3WayEnable);

fbValve(
    xEnable := (gxStart AND (DO_Pump1_T1_2 OR DO_Pump2_T1_2)) OR (gx3WayManual),
    iSV := SEL(gx3WayManual, giPID3WayTask, SV_3WayManualTask),
    iDlt := SEL(gx3WayManual, SV_3WayDelta, 0),
    (* Ход клапана задаётся с панели в СЕКУНДАХ, люфт - в МИЛЛИСЕКУНДАХ.
       Арифметику делаем в DINT(мс), в TIME переводим только результат *)
    tTotalTime := DINT_TO_TIME(INT_TO_DINT(SV_3WayTotalTime) * 1000),
    tLuftTime := DINT_TO_TIME(INT_TO_DINT(SV_3WayLuftTime)),
    xCloseOnDisable := gx3WayCloseWhenOff,
    xIsOpened := FALSE,
    xIsClosed := FALSE,
    xOpen := DO_3wayOpen,
    xClose := DO_3wayClose
);

(* Подпитка.
   Защита от переподпитки действует и в ручном режиме: RST стоит последним,
   поэтому при давлении выше SV_PresFilStop или аварии 33 клапан закрыт
   в любом режиме, даже если оператор держит ручную подпитку. *)
(* Авария 49 - датчик давления в системе показывает 0.0 бара (вероятно
   обрыв). Набирать воду по неработающему датчику нельзя: клапан открылся
   бы до аварии 34 по таймауту и залил систему. *)
SET(
    (gxFillManual OR (gxFillAuto AND AI_P_Set < SV_PresFilStart))
    AND NOT AM_ALARMS[49].Alarm,
    DO_ValveFill
);
RST(
    (NOT gxFillAuto AND NOT gxFillManual)
    OR (AI_P_Set > SV_PresFilStop)
    OR AM_ALARMS[33].Alarm (* Давление в системе выше максимума *),
    DO_ValveFill
);

(* Циркуляционные насосы *)
giWorkStages := 0;
FOR iCount := 0 TO c_HEATERS_IDX DO
    INC(arBurners[iCount].Stage1, giWorkStages);
    INC(arBurners[iCount].Stage2, giWorkStages);
END_FOR;

fbCirculation(
    ActiveStages := giWorkStages,
    ActivePupmp1 := gxEnablePump1 AND NOT (AM_ALARMS[21].Alarm OR AM_ALARMS[25].Alarm),
    ActivePupmp2 := gxEnablePump2 AND NOT (AM_ALARMS[22].Alarm OR AM_ALARMS[25].Alarm),
    ActivePupmp3 := gxEnablePump3 AND NOT (AM_ALARMS[23].Alarm OR AM_ALARMS[25].Alarm),
    ManualPupmp1 := gxManualPump1,
    ManualPupmp2 := gxManualPump2,
    ManualPupmp3 := gxManualPump3,
    Start := gxStart,
    StartPump1 := DO_Pump1,
    StartPump2 := DO_Pump2,
    StartPump3 := DO_Pump3
);

fbPumpsSO(
    EnableP1 := gxPump1_T1_Enable,
    EnableP2 := gxPump2_T1_Enable,
    ManualP1 := gxPump1_T1_Manual,
    ManualP2 := gxPump2_T1_Manual,
    AlarmP1 := AM_ALARMS[15].Alarm OR AM_ALARMS[25].Alarm,
    AlarmP2 := AM_ALARMS[16].Alarm OR AM_ALARMS[25].Alarm,
    RT := 1_728_000, (* 24 hours in 50ms increments *)
    PUMP1 := DO_Pump1_T1,
    PUMP2 := DO_Pump2_T1
);

fbPumpsToTO(
    EnableP1 := gxPump1_T1_2_Enable,
    EnableP2 := gxPump2_T1_2_Enable,
    ManualP1 := gxPump1_T1_2_Manual,
    ManualP2 := gxPump2_T1_2_Manual,
    AlarmP1 := AM_ALARMS[17].Alarm OR AM_ALARMS[25].Alarm,
    AlarmP2 := AM_ALARMS[18].Alarm OR AM_ALARMS[25].Alarm,
    RT := 1_728_000, (* 24 hours in 50ms increments *)
    PUMP1 := DO_Pump1_T1_2,
    PUMP2 := DO_Pump2_T1_2
);

fbPumpsFromTO(
    EnableP1 := gxPump1_T3_Enable,
    EnableP2 := gxPump2_T3_Enable,
    ManualP1 := gxPump1_T3_Manual,
    ManualP2 := gxPump2_T3_Manual,
    AlarmP1 := AM_ALARMS[19].Alarm,
    AlarmP2 := AM_ALARMS[20].Alarm,
    RT := 1_728_000, (* 24 hours in 50ms increments *)
    PUMP1 := DO_Pump1_T3,
    PUMP2 := DO_Pump2_T3
);
END_PROGRAM

PROGRAM PROCESS
VAR
  fbAmHasAlarm : FB_AM_HAS_ALARMS;
  fbAmSet : FB_AM_SET;
  fbAmReset : FB_AM_RESET;
  iAvailable : INT;
  iCount : INT;
  fbAMBuzzer : FB_AM_BUZZER;
  xBuzzerReset : BOOL;
  fbAMPack : FB_AM_PACK_ALARMS;
  fbAmHasAny : FB_AM_HAS_ALARMS;  (* Признак любой аварии для лампы *)
END_VAR
(* ==========================================================================
   PRG_PROCESS - обработка входов, аварий, состояний и моточасов.
   Карта аналоговых входов (модули Coolmay, R-регистры):
     R23700..R23702 - температура котлов 1..3 (Pt100, 0.1 C)
     R23703 - обратка отопления, R23705 - подача отопления
     R23704 - подача на котлы (коллектор), R23706/R23707 - теплообменник
     R23708 - температура наружного воздуха, R23709 - температура газа
     R23712..R23714 - давление котлов 1..3, R23715 - подача во внешнюю систему
     R23716 - обратка внешняя, R23717/R23718 - теплообменник
     R23719 - давление коллектора первичного контура (подпитка)
     D8032 - давление газа (встроенный вход модуля)
   Cor_* - поправки датчиков, задаются с панели.
   ========================================================================== *)
EI(TRUE);

AI_T_Heater1 := R23700 + Cor_T_Heater1;
AI_T_Heater2 := R23701 + Cor_T_Heater2;
AI_T_Heater3 := R23702 + Cor_T_Heater3;
AI_T_Colector := R23704 + Cor_T_Colector;
AI_T_SOFrom := R23703 + Cor_T_SOFrom;
AI_T_SOTo := R23705 + Cor_T_SOTo;
AI_T_GVSTo := R23706 + Cor_T_GVSTo;
AI_T_GVSFrom := R23707 + Cor_T_GVSFrom;
AI_T_Gaz := R23709 + Cor_T_Gaz;
AI_T_Weather := R23708 + Cor_T_Weather;

AI_P1 := F_SCALE(R23712, 0, 30000, 0, Max_P1, FALSE);
AI_P2 := F_SCALE(R23713, 0, 30000, 0, Max_P2, FALSE);
AI_P3 := F_SCALE(R23714, 0, 30000, 0, Max_P3, FALSE);
AI_P_SOTo := F_SCALE(R23715, 0, 30000, 0, Max_P_SOTo, FALSE);
AI_P_SOFrom := F_SCALE(R23716, 0, 30000, 0, Max_P_SOFrom, FALSE);
AI_P_GVSTo := F_SCALE(R23717, 0, 30000, 0, Max_P_GVSTo, FALSE);
AI_P_GVSFrom := F_SCALE(R23718, 0, 30000, 0, Max_P_GVSFrom, FALSE);
AI_P_Set := F_SCALE(R23719, 0, 30000, 0, Max_P_Set, FALSE);
AI_P_GAZ := F_SCALE(D8032, 0, 4030, 0, Max_P_GAZ, FALSE);

FAI_T_Heater1 := INT_TO_REAL(AI_T_Heater1) / 10.0;
FAI_T_Heater2 := INT_TO_REAL(AI_T_Heater2) / 10.0;
FAI_T_Heater3 := INT_TO_REAL(AI_T_Heater3) / 10.0;
FAI_T_Colector := INT_TO_REAL(AI_T_Colector) / 10.0;
FAI_T_SOFrom := INT_TO_REAL(AI_T_SOFrom) / 10.0;
FAI_T_SOTo := INT_TO_REAL(AI_T_SOTo) / 10.0;
FAI_T_GVSTo := INT_TO_REAL(AI_T_GVSTo) / 10.0;
FAI_T_GVSFrom := INT_TO_REAL(AI_T_GVSFrom) / 10.0;
FAI_T_Gaz := INT_TO_REAL(AI_T_Gaz) / 10.0;
FAI_T_Weather := INT_TO_REAL(AI_T_Weather) / 10.0;

FAI_P1 := INT_TO_REAL(AI_P1) / 10.0;
FAI_P2 := INT_TO_REAL(AI_P2) / 10.0;
FAI_P3 := INT_TO_REAL(AI_P3) / 10.0;
FAI_P_SOTo := INT_TO_REAL(AI_P_SOTo) / 10.0;
FAI_P_SOFrom := INT_TO_REAL(AI_P_SOFrom) / 10.0;
FAI_P_GVSTo := INT_TO_REAL(AI_P_GVSTo) / 10.0;
FAI_P_GVSFrom := INT_TO_REAL(AI_P_GVSFrom) / 10.0;
FAI_P_Set := INT_TO_REAL(AI_P_Set) / 10.0;
FAI_P_GAZ := INT_TO_REAL(AI_P_GAZ) / 10.0;

(* ОБРЫВ ДАТЧИКОВ ТЕМПЕРАТУРЫ. Модуль отдаёт ровно -1990 (-199.0 C) на
   разомкнутом Pt100, поэтому сравниваем с -1990 на равенство.
   Вход - сырые регистры АЦП R2370x, а не показания AI_T_*: в показаниях уже
   прибавлена поправка Cor_* с панели, и признак обрыва был бы искажён.
   Аварии 36/37/38 (котлы 1/2/3) идут в группы 1/2/3 - такой котёл
   выводится из каскада через arBurners[i].Error, как перегрев.
   Авария 39 (коллектор) и 43 (обратка ТО ГВС) дополнительно снимают
   ПИД каскада и ПИД 3-ходового клапана - см. PRG_MAIN.
   Аварии 40/41/42/44/45 - только сигнализация, в логике не участвуют. *)
fbAmSet(iNum := 36, xState := R23700 = -1990);   (* T котла 1 *)
fbAmSet(iNum := 37, xState := R23701 = -1990);   (* T котла 2 *)
fbAmSet(iNum := 38, xState := R23702 = -1990);   (* T котла 3 *)
fbAmSet(iNum := 39, xState := R23704 = -1990);   (* T коллектора *)
fbAmSet(iNum := 40, xState := R23703 = -1990);   (* T обратки отопления *)
fbAmSet(iNum := 41, xState := R23705 = -1990);   (* T подачи отопления *)
fbAmSet(iNum := 42, xState := R23706 = -1990);   (* T подачи ГВС *)
fbAmSet(iNum := 43, xState := R23707 = -1990);   (* T обратки ГВС *)
fbAmSet(iNum := 44, xState := R23709 = -1990);   (* T газа *)
fbAmSet(iNum := 45, xState := R23708 = -1990);   (* T улицы *)
(* НУЛЕВОЕ ДАВЛЕНИЕ (обрыв линии 4..20 мА или отказ датчика).
   На разомкнутой линии 4..20 мА модуль отдаёт ровно 0 (после F_SCALE это
   0.0 бара), поэтому сравниваем с 0 на равенство. Вход - сырые регистры
   R2371x, газ - встроенный вход D8032. Показание 2 отсчёта и выше означает
   живой датчик и тревоги не даёт: 2 отсчёта - это уже сигнал с датчика.
   Давление котла (46/47/48) идёт в группы 1/2/3 - котёл выходит из
   каскада, как при перегреве.
   Давление в системе (49), газа (50) и давлений отопления/ГВС (51..54) -
   группа 10, насосы они НЕ запрещают. По аварии 49 закрывается подпитка. *)
fbAmSet(iNum := 46, xState := R23712 = 0);   (* давление котла 1 *)
fbAmSet(iNum := 47, xState := R23713 = 0);   (* давление котла 2 *)
fbAmSet(iNum := 48, xState := R23714 = 0);   (* давление котла 3 *)
fbAmSet(iNum := 49, xState := R23719 = 0);   (* давление в системе *)
fbAmSet(iNum := 50, xState := D8032 = 0);    (* давление газа *)
fbAmSet(iNum := 51, xState := R23715 = 0);   (* давление подачи отопления *)
fbAmSet(iNum := 52, xState := R23716 = 0);   (* давление обратки отопления *)
fbAmSet(iNum := 53, xState := R23717 = 0);   (* давление подачи ГВС *)
fbAmSet(iNum := 54, xState := R23718 = 0);   (* давление обратки ГВС *)


T1_State := HEATER_STATE(arBurners[0]);
T2_State := HEATER_STATE(arBurners[1]);
T3_State := HEATER_STATE(arBurners[2]);

(* Состояние насоса для панели: 0 - выкл, 1 - работает, 2 - авария,
   4 - запрещён. Второй параметр - признак аварии насоса из менеджера тревог *)
Pump1_T1_State := PUMP_STATE(DO_Pump1_T1, AM_ALARMS[15].Alarm, gxPump1_T1_Enable);
Pump2_T1_State := PUMP_STATE(DO_Pump2_T1, AM_ALARMS[16].Alarm, gxPump2_T1_Enable);
Pump1_T1_2_State := PUMP_STATE(DO_Pump1_T1_2, AM_ALARMS[17].Alarm, gxPump1_T1_2_Enable);
Pump2_T1_2_State := PUMP_STATE(DO_Pump2_T1_2, AM_ALARMS[18].Alarm, gxPump2_T1_2_Enable);
Pump1_T3_State := PUMP_STATE(DO_Pump1_T3, AM_ALARMS[19].Alarm, gxPump1_T3_Enable);
Pump2_T3_State := PUMP_STATE(DO_Pump2_T3, AM_ALARMS[20].Alarm, gxPump2_T3_Enable);
Pump1_State := PUMP_STATE(DO_Pump1, AM_ALARMS[21].Alarm, gxEnablePump1);
Pump2_State := PUMP_STATE(DO_Pump2, AM_ALARMS[22].Alarm, gxEnablePump2);
Pump3_State := PUMP_STATE(DO_Pump3, AM_ALARMS[23].Alarm, gxEnablePump3);

IF AI_T_Weather <= SV_TWeather1 THEN
	giTSV := SV_TWater1;
ELSIF AI_T_Weather <= SV_TWeather2 THEN
	giTSV := F_SCALE(AI_T_Weather, SV_TWeather1, SV_TWeather2, SV_TWater1, SV_TWater2, FALSE);
ELSIF AI_T_Weather <= SV_TWeather3 THEN
	giTSV := F_SCALE(AI_T_Weather, SV_TWeather2, SV_TWeather3, SV_TWater2, SV_TWater3, FALSE);
ELSIF AI_T_Weather <= SV_TWeather4 THEN
	giTSV := F_SCALE(AI_T_Weather, SV_TWeather3, SV_TWeather4, SV_TWater3, SV_TWater4, FALSE);
ELSE
	giTSV := SV_TWater4;
END_IF;

fbAmSet(iNum := 0, xState := AI_T_Heater1 > SV_MaxTemperatureHeater);
fbAmSet(iNum := 1, xState := AI_P1 > SV_MaxPressure);
fbAmSet(iNum := 2, xState := AI_P1 < SV_MinPressure AND R23712 <> 0);
fbAmSet(iNum := 3, xState := DI_BurnAlarm1);
fbAmHasAlarm(iSeverity := c_AM_ERROR, iProcessNum := 1);
arBurners[0].Error := fbAmHasAlarm.Q;
arBurners[0].Manual := arBurners[0].Manual OR arBurners[0].ManualSecond;
arBurners[0].Work := DI_BurnWork1;
arBurners[0].Temperature := AI_T_Heater1;
arBurners[0].Pressure := AI_P1;
DO_Burn1Power := arBurners[0].Power;
DO_Burn1Stage1 := arBurners[0].Stage1;
DO_Burn1Stage2 := arBurners[0].Stage2;

fbAmSet(iNum := 5, xState := AI_T_Heater2 > SV_MaxTemperatureHeater);
fbAmSet(iNum := 6, xState := AI_P2 > SV_MaxPressure);
fbAmSet(iNum := 7, xState := AI_P2 < SV_MinPressure AND R23713 <> 0);
fbAmSet(iNum := 8, xState := DI_BurnAlarm2);
fbAmHasAlarm(iSeverity := c_AM_ERROR, iProcessNum := 2);
arBurners[1].Error := fbAmHasAlarm.Q;
arBurners[1].Manual := arBurners[1].Manual OR arBurners[1].ManualSecond;
arBurners[1].Work := DI_BurnWork2;
arBurners[1].Temperature := AI_T_Heater2;
arBurners[1].Pressure := AI_P2;
DO_Burn2Power := arBurners[1].Power;
DO_Burn2Stage1 := arBurners[1].Stage1;
DO_Burn2Stage2 := arBurners[1].Stage2;

fbAmSet(iNum := 10, xState := AI_T_Heater3 > SV_MaxTemperatureHeater);
fbAmSet(iNum := 11, xState := AI_P3 > SV_MaxPressure);
fbAmSet(iNum := 12, xState := AI_P3 < SV_MinPressure AND R23714 <> 0);
fbAmSet(iNum := 13, xState := DI_BurnAlarm3);
fbAmHasAlarm(iSeverity := c_AM_ERROR, iProcessNum := 3);
arBurners[2].Error := fbAmHasAlarm.Q;
arBurners[2].Manual := arBurners[2].Manual OR arBurners[2].ManualSecond;
arBurners[2].Work := DI_BurnWork3;
arBurners[2].Temperature := AI_T_Heater3;
arBurners[2].Pressure := AI_P3;
DO_Burn3Power := arBurners[2].Power;
DO_Burn3Stage1 := arBurners[2].Stage1;
DO_Burn3Stage2 := arBurners[2].Stage2;

(* DO_Pump1_T1 *)
fbAmSet(iNum := 15, xState := DO_Pump1_T1 AND NOT DI_Pump1_T1);
(* DO_Pump2_T1 *)
fbAmSet(iNum := 16, xState := DO_Pump2_T1 AND NOT DI_Pump2_T1);
(* DO_Pump1_T1_2 *)
fbAmSet(iNum := 17, xState := DO_Pump1_T1_2 AND NOT DI_Pump1_T1_2);
(* DO_Pump2_T1_2 *)
fbAmSet(iNum := 18, xState := DO_Pump2_T1_2 AND NOT DI_Pump2_T1_2);
(* DO_Pump1_T3 *)
fbAmSet(iNum := 19, xState := DO_Pump1_T3 AND NOT DI_Pump1_T3);
(* DO_Pump2_T3 *)
fbAmSet(iNum := 20, xState := DO_Pump2_T3 AND NOT DI_Pump2_T3);
(* DO_Pump1 *)
fbAmSet(iNum := 21, xState := DO_Pump1 AND NOT DI_Pump1);
(* DO_Pump2 *)
fbAmSet(iNum := 22, xState := DO_Pump2 AND NOT DI_Pump2);
(* DO_Pump3 *)
fbAmSet(iNum := 23, xState := DO_Pump3 AND NOT DI_Pump3);

iAvailable := 0;
FOR iCount := 0 TO c_HEATERS_IDX DO
    INC(
    	(arBurners[iCount].Auto OR arBurners[iCount].Manual)
    	AND NOT arBurners[iCount].Error
    	AND arBurners[iCount].Enable,
    	iAvailable
    );
END_FOR;

fbAmSet(iNum := 24, xState := AI_P_GAZ < SV_GasMinPressure);
(* 25 - давление в системе ниже минимального: запрет насосов.
   На 0.0 бара эта авария не срабатывает (там авария 49): обрыв датчика
   не должен останавливать насосы навсегда - иначе котельная не пустится. *)
fbAmSet(iNum := 25, xState := AI_P_Set < SV_SetMinPressure AND R23719 <> 0);
fbAmSet(iNum := 26, xState := NOT DI_EKM);
fbAmSet(iNum := 27, xState := NOT DI_ES);
fbAmSet(iNum := 28, xState := NOT DI_RKF);
fbAmSet(iNum := 29, xState := gxStart AND iAvailable = 0);
fbAmSet(iNum := 30, xState := gxNoSettings);

(* 31 - пуск котлов запрещён, пока не запущен хотя бы один насос.
   Проверяем ДО пуска (по gxStart), иначе первый цикл котлы включаются
   раньше насосов. Авария без защёлки и блокирующая (xLock = 1). *)
fbAmSet(iNum := 31, xState := gxStart AND NOT (DO_Pump1 OR DO_Pump2 OR DO_Pump3));

fbAmSet(iNum := 32, xState := AI_T_Colector > SV_MaxTemperatureColector);

fbAmSet(iNum := 33, xState := AI_P_Set > SV_MaxPressure);

OUT_T(DO_ValveFill, TC12, SV_MaxFillTime * 10);
fbAmSet(iNum := 34, xState := TS12);

fbAmSet(iNum := 35, xState := AI_T_GVSFrom > SV_3WayMaxTemperature);

(* 4, 9, 14 - термозащита котлов: авария, если пропал контакт (X035..X037).
   Номера взяты из резервных слотов групп котлов, поэтому тревога
   выводит из каскада только свой котёл, а упаковка для панели
   для панели остаётся сплошной: авария n уходит в бит M(530 + n), т.е. 534 / 539 / 544 *)
fbAmSet(iNum := 4, xState := NOT DI_BurnTherm1);
fbAmSet(iNum := 9, xState := NOT DI_BurnTherm2);
fbAmSet(iNum := 14, xState := NOT DI_BurnTherm3);

fbAMPack(DNUM := 530, PD := c_AM_PACK_M);

(* Наличие любой аварии берём у менеджера тревог, а не суммой упакованных битов:
   сумма 16-битная и могла переполниться в 0 *)
fbAmHasAny(iProcessNum := 0, iSeverity := 0);
gxHasalarm := fbAmHasAny.Q;
DO_AlarmLight := gxHasalarm;

(* Настройки считаются введёнными, если заполнены уставки и коэффициенты ПИД.
   R503 входит в блок параметров ПИД (R500..R528) и задаётся с панели:
   если он 0, значит коэффициенты регулятора не введены.
   Расчёт идёт ниже вызова fbAmSet(30) намеренно: авария реагирует
   с задержкой в один цикл, это допустимо. *)
gxNoSettings := (R503 = 0)
	OR (SV_TLimit = 0)
	OR (SV_MaxPressure = 0)
	OR (SV_MinPressure = 0)
	OR (SV_MaxTemperatureHeater = 0)
	OR (SV_TWeather1 = 0)
	OR (SV_TWeather2 = 0)
	OR (SV_TWeather3 = 0)
	OR (SV_TWeather4 = 0)
	OR (SV_TWater1 = 0)
	OR (SV_TWater2 = 0)
	OR (SV_TWater3 = 0)
	OR (SV_TWater4 = 0)
	OR (SV_GasMinPressure = 0)
	OR (SV_SetMinPressure = 0)
   OR (SV_3WayTempGVS = 0)
   OR (SV_HowOftenToCheck = 0)
   OR (SV_PresFilStart = 0)
   OR (SV_PresFilStop = 0)
   OR (SV_MaxFillTime = 0)
   OR (SV_3WayDelta = 0)
   OR (SV_3WayTotalTime = 0)
   OR (SV_3WayLuftTime = 0)
   OR (SV_3WayTempGVSDelta = 0)
   OR (SV_3WayManualTask = 0)
   OR (Max_P1 = 0)
	OR (Max_P2 = 0)
	OR (Max_P3 = 0)
	OR (Max_P_SOTo = 0)
	OR (Max_P_SOFrom = 0)
	OR (Max_P_GVSTo = 0)
	OR (Max_P_GVSFrom = 0)
	OR (Max_P_Set = 0)
	OR (Max_P_GAZ = 0)
   OR (SV_3WayMaxTemperature = 0)
   OR (SV_MaxTemperatureColector = 0)
    ;
(* Сброс аварий. IN - IN_OUT: блок держит импульс сброса 500 мс и сам гасит
   сигнал, поэтому отдельный RST не нужен. AutoReset не задаём: автосброс
   защёлкнутых аварий нужен только в особых случаях (например, однократный
   сбой связи, который слишком короткий, чтобы его заметила панель) *)
fbAmReset(IN := gxErrorReset);

(* Сирена. Блок сам защёлкивает Q, когда звуковых аварий стало больше,
   и снимает его по входу Reset, поэтому SET/RST не нужны.
   Reset - IN_OUT, в него можно передать только метку, поэтому кнопки сброса
   сводим в одну переменную *)
xBuzzerReset := gxResetAlarm OR gxErrorReset OR DI_AlarmReset;
fbAMBuzzer(Reset := xBuzzerReset, Q := DO_AlarmBuzzer);

(* Моточасы. У каждого счётчика свой флаг переполнения *)
HOUR(DO_Burn1Stage1, K32000, giHeater1Hours, gxWHOvfHeater1);
IF gxResetWHT1 THEN giHeater1Hours[0] := 0; giHeater1Hours[1] := 0; END_IF;
HOUR(DO_Burn2Stage1, K32000, giHeater2Hours, gxWHOvfHeater2);
IF gxResetWHT2 THEN giHeater2Hours[0] := 0; giHeater2Hours[1] := 0; END_IF;
HOUR(DO_Burn3Stage1, K32000, giHeater3Hours, gxWHOvfHeater3);
IF gxResetWHT3 THEN giHeater3Hours[0] := 0; giHeater3Hours[1] := 0; END_IF;
HOUR(DO_Pump1_T1, K32000, Pump1_T1_WH, gxWHOvfPump1_T1);
IF gxPump1_T1_WHReset THEN Pump1_T1_WH[0] := 0; Pump1_T1_WH[1] := 0; END_IF;
HOUR(DO_Pump2_T1, K32000, Pump2_T1_WH, gxWHOvfPump2_T1);
IF gxPump2_T1_WHReset THEN Pump2_T1_WH[0] := 0; Pump2_T1_WH[1] := 0; END_IF;
HOUR(DO_Pump1_T1_2, K32000, Pump1_T1_2_WH, gxWHOvfPump1_T1_2);
IF gxPump1_T1_2_WHReset THEN Pump1_T1_2_WH[0] := 0; Pump1_T1_2_WH[1] := 0; END_IF;
HOUR(DO_Pump2_T1_2, K32000, Pump2_T1_2_WH, gxWHOvfPump2_T1_2);
IF gxPump2_T1_2_WHReset THEN Pump2_T1_2_WH[0] := 0; Pump2_T1_2_WH[1] := 0; END_IF;
HOUR(DO_Pump1_T3, K32000, Pump1_T3_WH, gxWHOvfPump1_T3);
IF gxPump1_T3_WHReset THEN Pump1_T3_WH[0] := 0; Pump1_T3_WH[1] := 0; END_IF;
HOUR(DO_Pump2_T3, K32000, Pump2_T3_WH, gxWHOvfPump2_T3);
IF gxPump2_T3_WHReset THEN Pump2_T3_WH[0] := 0; Pump2_T3_WH[1] := 0; END_IF;
HOUR(DO_Pump1, K32000, Pump1_WH, gxWHOvfPump1);
IF gxPump1_WHReset THEN Pump1_WH[0] := 0; Pump1_WH[1] := 0; END_IF;
HOUR(DO_Pump2, K32000, Pump2_WH, gxWHOvfPump2);
IF gxPump2_WHReset THEN Pump2_WH[0] := 0; Pump2_WH[1] := 0; END_IF;
HOUR(DO_Pump3, K32000, Pump3_WH, gxWHOvfPump3);
IF gxPump3_WHReset THEN Pump3_WH[0] := 0; Pump3_WH[1] := 0; END_IF;
END_PROGRAM

PROGRAM INIT
VAR
  fbAmInit : FB_AM_INIT;
END_VAR
(* ==========================================================================
   PRG_INIT - инициализация контроллера.
   Вызывается ОДИН РАЗ по событию M8002 (начальный импульс), поэтому
   собственной защиты в коде нет.
   ========================================================================== *)
EI(TRUE);

(* --------------------------------------------------------------------------
   Параметры ПИД-регулятора КАСКАДА котлов - блок параметров R500..R528
   (29 слов, положение слова в блоке задано драйвером PID):
     R500 - время дискретизации (Ts), миллисекунды (1000 = 1 с)
     R501 - режим работы: 2#...0001 - обычный,
                  биты 4 (16) и 6 (64) включают автонастройку
     R502..R521 - коэффициенты P, I, D и остальные параметры контура.
                  Задаются оператором с панели и в программе НЕ
                  инициализируются (см. аварию 30 "нет настроек").
     R522 - верхний предел выхода, 600 = 100 %
     R523 - нижний предел выхода
     R525 - дельта автонастройки (5 = 0.5 бара)
     R526, R527 - пределы выхода во время автонастройки
     R528 - служебное слово блока ПИД
   -------------------------------------------------------------------------- *)
R500 := 1000; (* Период дискретизации ПИД 1 с (единица - мс) *)
R501 := 2#0000_0000_0000_0001; (* Heating mode *)
R522 := 600; (* Output max 100% *)
R523 := 0; (* Output min *)
R525 := 5; (* Delta for Autotune 0.5 bar *)
R526 := R522; (* Autotune output upper value *)
R527 := 0; (* Autotune output lower value *)

(* --------------------------------------------------------------------------
   Параметры ПИД-регулятора 3-ходового клапана ГВС - блок R600..R628.
   Смысл слов тот же, что и в блоке R500..R528. Выход 0..1000 (0..100.0 %).
   -------------------------------------------------------------------------- *)
R600 := 1000; (* Период дискретизации ПИД 1 с (единица - мс) *)
R601 := 2#0000_0000_0000_0001; (* Heating mode *)
R622 := 1000; (* Output max 100% *)
R623 := 0; (* Output min *)
R625 := 5; (* Delta for Autotune 0.5 bar *)
R626 := R622; (* Autotune output upper value *)
R627 := 0; (* Autotune output lower value *)

(* Количество аварий задаётся константой c_AM_ALARMS_NUM в GVL.csv (45, т.е.
   аварии 0..45). Раньше здесь было присваивание AM_ALARMS_NUM := 34 -
   границу массива AM_ALARMS в теле программы менять нельзя.
   AM_D_START - адрес начала энергонезависимой области менеджера тревог,
   задан настройкой библиотеки. *)

(* --------------------------------------------------------------------------
   Пределы шкал аналоговых входов (0.1 бара). Если оператор не ввёл значение
   (0), подставляется 16.0 бара.
   -------------------------------------------------------------------------- *)
MOV(Max_P2 = 0, 160, Max_P2);
MOV(Max_P3 = 0, 160, Max_P3);
MOV(Max_P1 = 0, 160, Max_P1);
MOV(Max_P_SOTo = 0, 160, Max_P_SOTo);
MOV(Max_P_SOFrom = 0, 160, Max_P_SOFrom);
MOV(Max_P_GVSTo = 0, 160, Max_P_GVSTo);
MOV(Max_P_GVSFrom = 0, 160, Max_P_GVSFrom);
MOV(Max_P_Set = 0, 160, Max_P_Set);
MOV(Max_P_GAZ = 0, 160, Max_P_GAZ);

(* --------------------------------------------------------------------------
   УСТАВКИ ПО УМОЛЧАНИЮ.
   Записываются в том же стиле, что и пределы шкал датчиков выше: 0 в уставке
   означает "не введена", и подставляется значение по умолчанию. Любое
   ненулевое значение, введённое оператором с панели, сохраняется при
   перезапуске (PRG_INIT работает по M8002, то есть при каждом включении).
   Поэтому 0 не является допустимым значением ни для одной из этих уставок.
   ВНИМАНИЕ: значения ориентировочные, перед пуском проверить на объекте.
   Давления - в 0.1 бара (как показания AI_P* ), SV_MaxFillTime - секунды.
   -------------------------------------------------------------------------- *)
(* Период проверки каскада, секунд (кратен дискретизации ПИД R500 = 1 с) *)
MOV(SV_HowOftenToCheck = 0, 30, SV_HowOftenToCheck);
(* Гистерезис добавления ступени, в единицах выхода ПИД (30 = 5 % от 600) *)
MOV(SV_StageHyst = 0, 50, SV_StageHyst); (* 5.0 % *)

(* Защиты по температуре, °C *)
MOV(SV_MaxTemperatureHeater = 0, 90, SV_MaxTemperatureHeater);
MOV(SV_MaxTemperatureColector = 0, 95, SV_MaxTemperatureColector);
MOV(SV_TLimit = 0, 5, SV_TLimit);

(* Защиты по давлению, 0.1 бара *)
MOV(SV_MaxPressure = 0, 40, SV_MaxPressure);
MOV(SV_MinPressure = 0, 10, SV_MinPressure);
MOV(SV_SetMinPressure = 0, 20, SV_SetMinPressure);
MOV(SV_PresFilStart = 0, 15, SV_PresFilStart);
MOV(SV_PresFilStop = 0, 25, SV_PresFilStop);
MOV(SV_GasMinPressure = 0, 30, SV_GasMinPressure); (* проверить по датчику газа *)
MOV(SV_MaxFillTime = 0, 300, SV_MaxFillTime);

(* Контур ГВС и 3-ходовой клапан *)
MOV(SV_3WayTempGVS = 0, 60, SV_3WayTempGVS);
MOV(SV_3WayTempGVSDelta = 0, 5, SV_3WayTempGVSDelta);
MOV(SV_3WayMaxTemperature = 0, 75, SV_3WayMaxTemperature);
MOV(SV_3WayDelta = 0, 50, SV_3WayDelta);
MOV(SV_3WayTotalTime = 0, 120, SV_3WayTotalTime); (* проверить по паспорту клапана *)
MOV(SV_3WayLuftTime = 0, 500, SV_3WayLuftTime);
MOV(SV_3WayManualTask = 0, 500, SV_3WayManualTask);

(* Кривая погодозависимости: улица -15/-5/+5/+15 °C -> подача 78/68/58/48 °C.
   Точки обязаны идти по возрастанию улицы, иначе F_SCALE посчитает неверно.
   Нулевых значений у точек быть не может: 0 там означает "не введена",
   по нему gxNoSettings включает аварию 30, а MOV вернёт значение по
   умолчанию. Поэтому значения по умолчанию выбраны ненулевыми. *)
MOV(SV_TWeather1 = 0, -15, SV_TWeather1);
MOV(SV_TWater1 = 0, 78, SV_TWater1);
MOV(SV_TWeather2 = 0, -5, SV_TWeather2);
MOV(SV_TWater2 = 0, 68, SV_TWater2);
MOV(SV_TWeather3 = 0, 5, SV_TWeather3);
MOV(SV_TWater3 = 0, 58, SV_TWater3);
MOV(SV_TWeather4 = 0, 15, SV_TWeather4);
MOV(SV_TWater4 = 0, 48, SV_TWater4);

(* Сторожевой таймер контроллера, 500 мс *)
D8000 := 500;

(* --------------------------------------------------------------------------
   Регистры R23500.. конфигурируют режим аналоговых каналов модулей:
   0 - вход подключён к Pt100, 1 - вход 4..20 мА.
   R23500..R23509 - 10 каналов Pt100,
   R23512..R23520 - 9 каналов 4..20 мА.
   -------------------------------------------------------------------------- *)
R23500 := 0;
R23501 := 0;
R23502 := 0;
R23503 := 0;
R23504 := 0;
R23505 := 0;
R23506 := 0;
R23507 := 0;
R23508 := 0;
R23509 := 0;
(* Входы 4-20мА *)
R23512 := 1;
R23513 := 1;
R23514 := 1;
R23515 := 1;
R23516 := 1;
R23517 := 1;
R23518 := 1;
R23519 := 1;
R23520 := 1;
(* Конфигурация быстрых входов/выходов ПЛК *)
R23940 := 0;
R23941 := 0;
R23942 := 1;
R23943 := 1;

(* ==========================================================================
   ОПИСАНИЕ АВАРИЙ. Все параметры указываются явно, чтобы вставка новой
   аварии в середину списка не меняла настройки последующих.
     iProcess - группа (1/2/3 - котёл 1/2/3, 7 - насосы, 10 - общие)
     iDelay - задержка срабатывания, единицы 100 мс (20 = 2 с)
     xLatch - защёлка (сброс только оператором)
     xBuzzer - вывод на сирену
     xLock - блокировка работы каскада (группа -> fbAmBlock)
   ========================================================================== *)
fbAmInit.iSeverity := c_AM_ERROR;

(* --- Котёл 1 --------------------------------------------------------- *)
(* 0 - перегрев котла: котёл выводится из каскада *)
fbAmInit(iNum := 0, iProcess := 1, iDelay := 0,
         xLatch := 1, xBuzzer := 1, xLock := 0);
(* 1 - давление в котле выше SV_MaxPressure *)
fbAmInit(iNum := 1, iProcess := 1, iDelay := 0,
         xLatch := 0, xBuzzer := 1, xLock := 0);
(* 2 - давление в котле ниже SV_MinPressure *)
fbAmInit(iNum := 2, iProcess := 1, iDelay := 0,
         xLatch := 0, xBuzzer := 1, xLock := 0);
(* 3 - авария горелки (DI_BurnAlarm1) *)
fbAmInit(iNum := 3, iProcess := 1, iDelay := 0,
         xLatch := 1, xBuzzer := 1, xLock := 0);
(* 4 - котёл 1: пропал контакт термозащиты (X035) *)
fbAmInit(iNum := 4, iProcess := 1, iDelay := 20,
         xLatch := 1, xBuzzer := 1, xLock := 0);

(* --- Котёл 2 --------------------------------------------------------- *)
(* 5 - перегрев котла *)
fbAmInit(iNum := 5, iProcess := 2, iDelay := 0,
         xLatch := 1, xBuzzer := 1, xLock := 0);
(* 6 - давление в котле выше SV_MaxPressure *)
fbAmInit(iNum := 6, iProcess := 2, iDelay := 0,
         xLatch := 0, xBuzzer := 1, xLock := 0);
(* 7 - давление в котле ниже SV_MinPressure *)
fbAmInit(iNum := 7, iProcess := 2, iDelay := 0,
         xLatch := 0, xBuzzer := 1, xLock := 0);
(* 8 - авария горелки (DI_BurnAlarm2) *)
fbAmInit(iNum := 8, iProcess := 2, iDelay := 0,
         xLatch := 1, xBuzzer := 1, xLock := 0);
(* 9 - котёл 2: пропал контакт термозащиты (X036) *)
fbAmInit(iNum := 9, iProcess := 2, iDelay := 20,
         xLatch := 1, xBuzzer := 1, xLock := 0);

(* --- Котёл 3 --------------------------------------------------------- *)
(* 10 - перегрев котла *)
fbAmInit(iNum := 10, iProcess := 3, iDelay := 0,
         xLatch := 1, xBuzzer := 1, xLock := 0);
(* 11 - давление в котле выше SV_MaxPressure *)
fbAmInit(iNum := 11, iProcess := 3, iDelay := 0,
         xLatch := 0, xBuzzer := 1, xLock := 0);
(* 12 - давление в котле ниже SV_MinPressure *)
fbAmInit(iNum := 12, iProcess := 3, iDelay := 0,
         xLatch := 0, xBuzzer := 1, xLock := 0);
(* 13 - авария горелки (DI_BurnAlarm3) *)
fbAmInit(iNum := 13, iProcess := 3, iDelay := 0,
         xLatch := 1, xBuzzer := 1, xLock := 0);
(* 14 - котёл 3: пропал контакт термозащиты (X037) *)
fbAmInit(iNum := 14, iProcess := 3, iDelay := 20,
         xLatch := 1, xBuzzer := 1, xLock := 0);

(* --- Насосы: нет подтверждения работы (2 с) -------------------------- *)
(* 15 - насос 1 контура Т1 *)
fbAmInit(iNum := 15, iProcess := 7, iDelay := 20,
         xLatch := 1, xBuzzer := 1, xLock := 0);
(* 16 - насос 2 контура Т1 *)
fbAmInit(iNum := 16, iProcess := 7, iDelay := 20,
         xLatch := 1, xBuzzer := 1, xLock := 0);
(* 17 - насос 1 контура Т1.2 *)
fbAmInit(iNum := 17, iProcess := 7, iDelay := 20,
         xLatch := 1, xBuzzer := 1, xLock := 0);
(* 18 - насос 2 контура Т1.2 *)
fbAmInit(iNum := 18, iProcess := 7, iDelay := 20,
         xLatch := 1, xBuzzer := 1, xLock := 0);
(* 19 - насос 1 контура Т3 *)
fbAmInit(iNum := 19, iProcess := 7, iDelay := 20,
         xLatch := 1, xBuzzer := 1, xLock := 0);
(* 20 - насос 2 контура Т3 *)
fbAmInit(iNum := 20, iProcess := 7, iDelay := 20,
         xLatch := 1, xBuzzer := 1, xLock := 0);
(* 21 - насос 1 малого котлового контура *)
fbAmInit(iNum := 21, iProcess := 7, iDelay := 20,
         xLatch := 1, xBuzzer := 1, xLock := 0);
(* 22 - насос 2 малого котлового контура *)
fbAmInit(iNum := 22, iProcess := 7, iDelay := 20,
         xLatch := 1, xBuzzer := 1, xLock := 0);
(* 23 - насос 3 малого котлового контура *)
fbAmInit(iNum := 23, iProcess := 7, iDelay := 20,
         xLatch := 1, xBuzzer := 1, xLock := 0);

(* --- Общие аварии ---------------------------------------------------- *)
(* 24 - давление газа ниже SV_GasMinPressure, блокирует *)
fbAmInit(iNum := 24, iProcess := 10, iDelay := 0,
         xLatch := 0, xBuzzer := 0, xLock := 1);
(* 25 - давление подпитки ниже SV_SetMinPressure (запрет насосов) *)
fbAmInit(iNum := 25, iProcess := 10, iDelay := 0,
         xLatch := 0, xBuzzer := 0, xLock := 0);
(* 26 - нет питания ЭКМ *)
fbAmInit(iNum := 26, iProcess := 10, iDelay := 0,
         xLatch := 1, xBuzzer := 1, xLock := 1);
(* 27 - нет питания аварийной кнопки (ES) *)
fbAmInit(iNum := 27, iProcess := 10, iDelay := 0,
         xLatch := 0, xBuzzer := 1, xLock := 1);
(* 28 - нет питания РКФ *)
fbAmInit(iNum := 28, iProcess := 10, iDelay := 0,
         xLatch := 0, xBuzzer := 0, xLock := 1);
(* 29 - нет ни одного доступного котла при пуске *)
fbAmInit(iNum := 29, iProcess := 10, iDelay := 0,
         xLatch := 0, xBuzzer := 1, xLock := 1);
(* 30 - не введены настройки (gxNoSettings), блокирует *)
fbAmInit(iNum := 30, iProcess := 10, iDelay := 0,
         xLatch := 0, xBuzzer := 0, xLock := 1);
(* 31 - ни один насос не запущен, пуск котлов запрещён.
       Без защёлки, т.к. снимается сама при пуске насоса,
       но блокирующая - иначе ошибку не видно. *)
fbAmInit(iNum := 31, iProcess := 10, iDelay := 20,
         xLatch := 0, xBuzzer := 0, xLock := 1);
(* 32 - перегрев коллектора. Мягкий лимит: снимает работу ПИД,
       но не блокирует каскад *)
fbAmInit(iNum := 32, iProcess := 10, iDelay := 20,
         xLatch := 0, xBuzzer := 0, xLock := 0);
(* 33 - давление в системе выше SV_MaxPressure (запрет подпитки) *)
fbAmInit(iNum := 33, iProcess := 10, iDelay := 20,
         xLatch := 0, xBuzzer := 0, xLock := 0);
(* 34 - подпитка не набирает воду за SV_MaxFillTime *)
fbAmInit(iNum := 34, iProcess := 10, iDelay := 0,
         xLatch := 0, xBuzzer := 0, xLock := 0);
(* 35 - температура ГВС выше SV_3WayMaxTemperature *)
fbAmInit(iNum := 35, iProcess := 10, iDelay := 0,
         xLatch := 0, xBuzzer := 0, xLock := 0);

(* --- Обрыв датчиков температуры --------------------------------------
   Модуль отдаёт ровно -1990 (-199.0 C) на разомкнутом Pt100. Условия
   (сырой регистр АЦП = -1990) выставляются в PRG_PROCESS.
   Обрыв датчика котла (36/37/38) в группах 1/2/3 выводит из каскада
   только свой котёл - через arBurners[i].Error. Остальные датчики котёл
   не останавливают:
     39 - коллектор: вход ПИД каскада, снимает регулятор,
     43 - обратка ТО ГВС: вход ПИД 3-ходового клапана, снимает регулятор,
     40/41/42/44/45 - только сигнализация.
   Защёлки нет: после ремонта датчика авария уходит сама.
   У датчиков ПИД (39, 43) задержки нет: регулятор нужно снимать сразу,
   иначе он успевает отработать по -199 C. Остальным датчикам 2 с, чтобы
   короткий сбой линии не ронял котёл. *)
(* 36 - обрыв датчика температуры котла 1 *)
fbAmInit(iNum := 36, iProcess := 1, iDelay := 20,
         xLatch := 0, xBuzzer := 1, xLock := 0);
(* 37 - обрыв датчика температуры котла 2 *)
fbAmInit(iNum := 37, iProcess := 2, iDelay := 20,
         xLatch := 0, xBuzzer := 1, xLock := 0);
(* 38 - обрыв датчика температуры котла 3 *)
fbAmInit(iNum := 38, iProcess := 3, iDelay := 20,
         xLatch := 0, xBuzzer := 1, xLock := 0);
(* 39 - обрыв датчика температуры коллектора (обратка от котлов): вход ПИД, без задержки *)
fbAmInit(iNum := 39, iProcess := 10, iDelay := 0,
         xLatch := 0, xBuzzer := 1, xLock := 0);
(* 40 - обрыв датчика температуры обратки отопления *)
fbAmInit(iNum := 40, iProcess := 10, iDelay := 20,
         xLatch := 0, xBuzzer := 1, xLock := 0);
(* 41 - обрыв датчика температуры подачи отопления *)
fbAmInit(iNum := 41, iProcess := 10, iDelay := 20,
         xLatch := 0, xBuzzer := 1, xLock := 0);
(* 42 - обрыв датчика температуры подачи на теплообменник ГВС *)
fbAmInit(iNum := 42, iProcess := 10, iDelay := 20,
         xLatch := 0, xBuzzer := 1, xLock := 0);
(* 43 - обрыв датчика температуры обратки с теплообменника ГВС: вход ПИД, без задержки *)
fbAmInit(iNum := 43, iProcess := 10, iDelay := 0,
         xLatch := 0, xBuzzer := 1, xLock := 0);
(* 44 - обрыв датчика температуры газа *)
fbAmInit(iNum := 44, iProcess := 10, iDelay := 20,
         xLatch := 0, xBuzzer := 1, xLock := 0);
(* 45 - обрыв датчика температуры наружного воздуха *)
fbAmInit(iNum := 45, iProcess := 10, iDelay := 20,
         xLatch := 0, xBuzzer := 1, xLock := 0);
(* --- Нулевое давление (обрыв линии 4..20 мА или отказ датчика) --------------
   На разомкнутой линии 4..20 мА модуль отдаёт 0, после F_SCALE это 0.0 бара.
   От настоящего нуля давления такой же код отличить нельзя, поэтому тревога
   и названа "вероятно обрыв". Сравнение - сырой регистр АЦП = 0 (0.0 бар).
   Задержки нет: 0.0 бара - состояние не мгновенное, а отказное.
   Обрыв датчика давления котла (46/47/48) идёт в группы 1/2/3 и выводит из
   каскада только свой котёл - как перегрев и обрыв датчика температуры.
   Остальные (49..54) котёл не останавливают и НЕ запрещают насосы:
     49 - давление в системе (подпитка), клапан подпитки при этом закрыт,
     50 - давление газа, каскад дополнительно блокирует авария 24,
     51/52/53/54 - давления отопления и ГВС, только сигнализация.
   Защёлки нет. *)
(* 46 - давление котла 1 равно 0.0 бара (вероятно обрыв датчика) *)
fbAmInit(iNum := 46, iProcess := 1, iDelay := 0,
         xLatch := 0, xBuzzer := 1, xLock := 0);
(* 47 - давление котла 2 равно 0.0 бара (вероятно обрыв датчика) *)
fbAmInit(iNum := 47, iProcess := 2, iDelay := 0,
         xLatch := 0, xBuzzer := 1, xLock := 0);
(* 48 - давление котла 3 равно 0.0 бара (вероятно обрыв датчика) *)
fbAmInit(iNum := 48, iProcess := 3, iDelay := 0,
         xLatch := 0, xBuzzer := 1, xLock := 0);
(* 49 - давление в системе 0.0 бара (вероятно обрыв датчика) *)
fbAmInit(iNum := 49, iProcess := 10, iDelay := 0,
         xLatch := 0, xBuzzer := 1, xLock := 0);
(* 50 - давление газа 0.0 бара (вероятно обрыв датчика) *)
fbAmInit(iNum := 50, iProcess := 10, iDelay := 0,
         xLatch := 0, xBuzzer := 1, xLock := 0);
(* 51 - давление подачи отопления 0.0 бара (вероятно обрыв датчика) *)
fbAmInit(iNum := 51, iProcess := 10, iDelay := 0,
         xLatch := 0, xBuzzer := 1, xLock := 0);
(* 52 - давление обратки отопления 0.0 бара (вероятно обрыв датчика) *)
fbAmInit(iNum := 52, iProcess := 10, iDelay := 0,
         xLatch := 0, xBuzzer := 1, xLock := 0);
(* 53 - давление подачи ГВС 0.0 бара (вероятно обрыв датчика) *)
fbAmInit(iNum := 53, iProcess := 10, iDelay := 0,
         xLatch := 0, xBuzzer := 1, xLock := 0);
(* 54 - давление обратки ГВС 0.0 бара (вероятно обрыв датчика) *)
fbAmInit(iNum := 54, iProcess := 10, iDelay := 0,
         xLatch := 0, xBuzzer := 1, xLock := 0);
END_PROGRAM

FUNCTION REVERSE
VAR_INPUT
  CUR : INT;
  MAX : INT;  (* Максимальный индекс. Например 0..5 значит 5 *)
END_VAR
REVERSE := ABS(CUR - MAX);
END_FUNCTION

FUNCTION_BLOCK Circulation
VAR_INPUT
  ActiveStages : INT;
  ActivePupmp1 : BOOL;
  ActivePupmp2 : BOOL;
  ActivePupmp3 : BOOL;
  ManualPupmp1 : BOOL;
  ManualPupmp2 : BOOL;
  ManualPupmp3 : BOOL;
  TimeinWork : INT;
  Start : BOOL;
END_VAR
VAR_OUTPUT
  StartPump1 : BOOL;
  StartPump2 : BOOL;
  StartPump3 : BOOL;
END_VAR
VAR
  Times : ARRAY [0..2] OF INT;
  Active : ARRAY [0..2] OF INT;
  NewTime : TON;
  NPump : INT;
  Pumps : ARRAY [0..2] OF PUMP;
  NambPump : INT;
  Order : INT;
  Restart : BOOL;
  ChangeN : INT;
  ChangeN2 : INT;
END_VAR
(* ==========================================================================
FB_Circulation - выбор работающих циркуляционных насосов малого контура.
Число насосов зависит от количества включённых ступеней котлов,
ведущий насос меняется раз в 24 часа для выравнивания моточасов.
Ручной пуск насоса имеет приоритет.
========================================================================== *)
CASE  ActiveStages  OF
	0..2 :
		NambPump := 1;
	3..4 :
		NambPump := 2;
	5..6 :
		NambPump := 3;			
END_CASE;

ChangeN := bool_to_int( ActivePupmp1 ) + bool_to_int( ActivePupmp2 ) + bool_to_int( ActivePupmp3 ) + bool_to_int( Start )
		+ bool_to_int( ManualPupmp1 ) + bool_to_int(ManualPupmp2 ) + bool_to_int( ManualPupmp3 ) + NambPump;
		
IF ChangeN <> ChangeN2 THEN
	Restart := TRUE;
	ChangeN2 := ChangeN;
END_IF;			 


Pumps[0].Evailable := ActivePupmp1;
Pumps[1].Evailable := ActivePupmp2;
Pumps[2].Evailable := ActivePupmp3;


(* Ведущий насос меняется раз в 24 часа. PT задаётся в TIME (мс),
поэтому считаем в DINT и только результат переводим в TIME *)
NewTime(IN := (Start AND NOT NewTime.Q), PT := DINT_TO_TIME(INT_TO_DINT(24) * 3600 * 1000));


IF NewTime.Q THEN
	Order := Order + 1;
	IF Order > 2 THEN
		Order := 0;
	END_IF;
	Restart	:= TRUE;	
END_IF;

IF Restart THEN 	
	
	FOR NPump := 0 TO 2 DO
			Pumps[NPump].Start := FALSE;			
	END_FOR;
	
	Pumps[0].Start := ManualPupmp1 AND Pumps[0].Evailable;
	Pumps[1].Start := ManualPupmp2 AND Pumps[1].Evailable;
	Pumps[2].Start := ManualPupmp3 AND Pumps[2].Evailable;
	
	FOR NPump := 0 TO 2 DO	
		IF Pumps[NPump].Start THEN
			NambPump := NambPump - 1;
		END_IF;			
	END_FOR;
	
	(* NambPump - сколько насосов ещё нужно запустить после ручных.
	Раньше здесь стояло NPump, а после цикла FOR эта переменная всегда 3 *)
	IF NambPump > 0 THEN
		FOR NPump := Order  TO 2 DO
			IF (Pumps[NPump].Evailable = TRUE) AND NOT (Pumps[NPump].Start = TRUE) AND NambPump > 0 THEN
				Pumps[NPump].Start := TRUE;
				NambPump := NambPump - 1;
			END_IF;	
			
			IF NambPump < 1 THEN
				EXIT;
			END_IF;			
		END_FOR;
		
		FOR NPump := 0 TO 2 DO
			IF (Pumps[NPump].Evailable = TRUE) AND NOT (Pumps[NPump].Start = TRUE) AND NambPump > 0 THEN
				Pumps[NPump].Start := TRUE;
				NambPump := NambPump - 1;
			END_IF;	
			IF NambPump < 1 THEN
				EXIT;
			END_IF;			
		END_FOR;
	END_IF;	
	Restart := FALSE;
END_IF;

IF NOT Start THEN
	Pumps[0].Start := FALSE;
	Pumps[1].Start := FALSE;
	Pumps[2].Start := FALSE;
END_IF;

StartPump1 := Pumps[0].Start AND Pumps[0].Evailable;
StartPump2 := Pumps[1].Start AND Pumps[1].Evailable;
StartPump3 := Pumps[2].Start AND Pumps[2].Evailable;
END_FUNCTION_BLOCK

FUNCTION HEATER_STATE
VAR_INPUT
  BURNER : BURNER;
END_VAR
HEATER_STATE := 0;

IF NOT BURNER.Power THEN		
    RETURN;
END_IF;

HEATER_STATE := 1;

IF BURNER.Stage1 THEN
	HEATER_STATE := 2;
END_IF;

IF BURNER.Stage2 THEN
	HEATER_STATE := 3;
END_IF;
END_FUNCTION

FUNCTION PUMP_STATE
VAR_INPUT
  PumpDO : BOOL;
  PumpAlarm : BOOL;
  PumpEnable : BOOL;
END_VAR
PUMP_STATE := SEL(
	PumpAlarm, 
	SEL(PumpEnable, 4, SEL(PumpDO, 0, 1)), 
	2
);
END_FUNCTION

FUNCTION_BLOCK PUMPS
VAR_INPUT
  EnableP1 : BOOL;
  EnableP2 : BOOL;
  ManualP1 : BOOL;
  ManualP2 : BOOL;
  AlarmP1 : BOOL;
  AlarmP2 : BOOL;
  RT : DWORD;
END_VAR
VAR_OUTPUT
  PUMP1 : BOOL;
  PUMP2 : BOOL;
END_VAR
VAR
  fbBlink : FB_TCO_50_BLINK;
  xBlink : BOOL;
END_VAR
(* ==========================================================================
   FB_PUMPS - два насоса контура Т1/Т1.2, работают по очереди (раз в RT).
   Насосы пускаются отдельно от котлов и не зависят от gxStart.
   Авария или запрет насоса снимает его выход и передаёт работу второму.
   ========================================================================== *)
fbBlink(xIn := TRUE, dwTimeLow := RT, dwTimeHigh := RT, xQ := xBlink);
PUMP1 := NOT AlarmP1 AND EnableP1 AND (ManualP1 OR xBlink OR (NOT xBlink AND (AlarmP2 OR NOT EnableP2)));
PUMP2 := NOT AlarmP2 AND EnableP2 AND (ManualP2 OR NOT xBlink OR (xBlink AND (AlarmP1 OR NOT EnableP1)));
END_FUNCTION_BLOCK
